    HMI_Message_Request : ARRAY[0..121] OF BOOL;  (* #HMI メッセージ表示要求; [0] 未使用; [1] 【Y616】A(左側) 供給スライド戻 異常表示; [2] 【Y617】A(左側) 供給スライド行 異常表示; [3] 【Y618】A(左側) 供給ピックアップ戻 異常表示; [4] 【Y619】A(左側) 供給ピックアップ行 異常表示; [5] 【Y620】A(左側) 供給チャック閉 戻 異常表示; [6] 【Y621】A(左側) 供給チャック開 行 異常表示; [7] 【Y622】B(右側) 供給スライド戻 異常表示; [8] 【Y623】B(右側) 供給スライド行 異常表示; [9] 【Y624】B(右側) 供給ピックアップ戻 異常表示; [10] 【Y625】B(右側) 供給ピックアップ行 異常表示; [11] 【Y626】B(右側) 供給チャック閉 戻 異常表示; [12] 【Y627】B(右側) 供給チャック開 行 異常表示; [13] 【Y700】A(左側) 高さ検査押え戻 異常表示; [14] 【Y701】A(左側) 高さ検査押え行 異常表示; [15] 【Y702】A(左側) 高さ検査持上戻 異常表示; [16] 【Y703】A(左側) 高さ検査持上行 異常表示; [17] 【Y704】A(左側) NG1ピックアップ戻 異常表示; [18] 【Y705】A(左側) NG1ピックアップ 行 異常表示; [19] 【Y706】A(左側) NG1チャック戻 異常表示; [20] 【Y707】A(左側) NG1チャック行 異常表示; [21] 【Y708】A(左側)ST4 反転1チャック閉 異常表示; [22] 【Y709】A(左側)ST4 反転1チャック開 異常表示; [23] 【Y710】A(左側)ST4 反転1ピックアップ戻 異常表示; [24] 【Y711】A(左側)ST4 反転1ピックアップ行 異常表示; [25] 【Y712】A(左側)ST6 反転2チャック閉 戻 異常表示; [26] 【Y713】A(左側)ST6 反転2チャック開 行 異常表示; [27] 【Y714】A(左側)ST6 反転2ピックアップ戻 異常表示; [28] 【Y715】A(左側)ST6 反転2ピックアップ行 異常表示; [29] 【Y716】A(左側) 排出チャック閉 戻 異常表示; [30] 【Y717】A(左側) 排出チャック開 行 異常表示; [31] 【Y718】A(左側) 排出フォルダ送り戻 異常表示; [32] 【Y719】A(左側) 排出フォルダ送り行 異常表示; [33] A(左側) 位置1ストッパー戻 異常表示; [34] 【Y720】A(左側) 位置1ストッパー 行 異常表示; [35] 【Y721】A(左側) 位置2ストッパー 異常表示; [36] 【Y721】A(左側) 位置2ストッパー 異常表示; [37] 【Y722】A(左側) 位置3ストッパー戻 異常表示; [38] 【Y722】A(左側) 位置3ストッパー行 異常表示; [39] Output_A_Error_M[33] 異常表示; [40] 【Y723】A(左側) 位置4ストッパー行 異常表示; [41] 【Y724】A(左側) 位置5ストッパー戻 異常表示; [42] 【Y724】A(左側) 位置5ストッパー行 異常表示; [43] 【Y725】A(左側) 位置6ストッパー戻 異常表示; [44] 【Y725】A(左側) 位置6ストッパー行 異常表示; [45] 【Y726】A(左側) ストックフォルダターン戻 異常表示; [46] 【Y727】A(左側) ストックフォルダターン行 異常表示; [47] 【Y728】A(左側) NG1仕分け 戻 異常表示; [48] 【Y729】A(左側) NG1仕分け 行 異常表示; [49] 【Y800】B(右側) 高さ検査押え戻 異常表示; [50] 【Y801】B(右側) 高さ検査押え行 異常表示; [51] 【Y802】B(右側) 高さ検査持上戻 異常表示; [52] 【Y803】B(右側) 高さ検査持上行 異常表示; [53] 【Y804】B(右側) NG1ピックアップ戻 異常表示; [54] 【Y805】B(右側) NG1ピックアップ 行 異常表示; [55] 【Y806】B(右側) NG1チャック戻 異常表示; [56] 【Y807】B(右側) NG1チャック行 異常表示; [57] 【Y808】B(右側)ST4 反転1チャック閉 戻 異常表示; [58] 【Y809】B(右側)ST4 反転1チャック開 戻 異常表示; [59] 【Y810】B(右側)ST4 反転1ピックアップ戻 異常表示; [60] 【Y811】B(右側)ST4 反転1ピックアップ行 異常表示; [61] 【Y812】B(右側)ST6 反転2チャック閉 戻 異常表示; [62] 【Y813】B(右側)ST6 反転2チャック開 行 異常表示; [63] 【Y814】B(右側)ST6 反転2ピックアップ戻 異常表示; [64] 【Y815】B(右側)ST6 反転2ピックアップ行 異常表示; [65] 【Y816】B(右側) 排出チャック閉 戻 異常表示; [66] 【Y817】B(右側) 排出チャック開 行 異常表示; [67] 【Y818】B(右側) 排出フォルダ送り戻 異常表示; [68] 【Y819】B(右側) 排出フォルダ送り行 異常表示; [69] 【Y820】B(右側) 位置1ストッパー 戻 異常表示; [70] 【Y820】B(右側) 位置1ストッパー 行 異常表示; [71] 【Y821】B(右側) 位置2ストッパー戻 異常表示; [72] 【Y821】B(右側) 位置2ストッパー行 異常表示; [73] 【Y822】B(右側) 位置3ストッパー戻 異常表示; [74] 【Y822】B(右側) 位置3ストッパー行 異常表示; [75] 【Y823】B(右側) 位置4ストッパー戻 異常表示; [76] 【Y823】B(右側) 位置4ストッパー行 異常表示; [77] 【Y824】B(右側) 位置5ストッパー戻 異常表示; [78] 【Y824】B(右側) 位置5ストッパー行 異常表示; [79] 【Y825】B(右側) 位置6ストッパー戻 異常表示; [80] 【Y825】B(右側) 位置6ストッパー行 異常表示; [81] 【Y826】B(右側) ストックフォルダターン戻 異常表示; [82] 【Y827】B(右側) ストックフォルダターン行 異常表示; [83] 【Y828】B(右側) NG1仕分け 戻 異常表示; [84] 【Y829】B(右側) NG1仕分け 行 異常表示; [85] 【Y1200】空コンテナ送り 戻 異常表示; [86] 【Y1201】空コンテナ送り 行 異常表示; [87] 【Y1202】段バラシ爪 戻 異常表示; [88] 【Y1203】段バラシ爪 行 異常表示; [89] 【Y1204】コンテナ排出 戻 異常表示; [90] 【Y1205】コンテナ排出 行 異常表示; [91] Output_Share_Error_M[7] 異常表示; [92] 【Y1207】箱入れチャック 行 異常表示; [93] 【Y1208】コンテナ仕分けストッパー 戻 異常表示; [94] 【Y1209】コンテナ仕分けストッパー 行 異常表示; [95] 【Y1210】コンテナ仕分け送り 戻 異常表示; [96] Output_Share_Error_M[12] 異常表示; [97] 【Y1300】A(左側) コンベア受渡送り戻 異常表示; [98] 【Y1301】A(左側) コンベア受渡送り行 異常表示; [99] 【Y1302】B(右側) コンベア受渡送り戻 異常表示; [100] 【Y1303】B(右側) コンベア受渡送り行 異常表示; [101] ST1 搬送ワーク不一致; [102] ST2 搬送ワーク不一致; [103] ST3 搬送ワーク不一致; [104] ST4 搬送ワーク不一致; [105] ST5 搬送ワーク不一致; [106] ST6 搬送ワーク不一致; [107] ST7 搬送ワーク不一致; [108] A(左側) ST1 FH測定時間超過; [109] A(左側) ST1 FH異常; [110] A(左側) ST5 FH異常; [111] B(右側) ST1 FH異常; [112] B(右側) ST5 FH異常; [113] A(左側) ST1 FH判定OK; [114] A(左側) ST1 FH判定NG1; [115] A(左側) ST1 FH判定NG2; [116] A(左側) ST1 検査前ワーク不一致; [117] A(左側) ST5 FH測定時間超過; [118] A(左側) ST5 FH判定OK; [119] A(左側) ST5 FH判定NG1; [120] A(左側) ST5 FH判定NG2; [121] A(左側) ST5 検査前ワーク不一致 *)
END_VAR

PROGRAM ModeManagement_モード管理
VAR
    Setting_M : BOOL;
    Manual_M : BOOL;
    Auto_M : BOOL;
    Dummy_M : BOOL;
    Inital_M : BOOL;
    Output_Error_M : ARRAY[0..99] OF Bool;
    Index_Error_001 : DINT;
    Index_B_001 : DINT;
    Index_Share_001 : DINT;
    Error_TON : ARRAY[0..99] OF TON;  (* [2] A(左側) ST1 測定タイムアウト; [4] A(左側) ST5 測定タイムアウト *)
    Error_TOF : ARRAY[0..99] OF TOF;
    AutoMode_A_M : ARRAY[0..99] OF Bool;
    ６ : DINT;
    ST4_A_Rev_01_Origin_M : ARRAY[0..99] OF Bool;  (* A(左側) ST4 反転1 原点復帰工程; [1] A(左側) ST4 反転1 原点復帰開始; [2] A(左側) ST4 反転1 原点復帰中; [3] A(左側) ST4 反転1 ピックアップ戻; [4] A(左側) ST4 反転1 モータ原点復帰開始; [5] A(左側) ST4 反転1 ピックアップ行; [6] A(左側) ST4 反転1 チャック閉; [7] A(左側) ST4 反転1 原点復帰完了（ワーク無） *)
    ST4_A_Rev_01_OriginDone : BOOL;  (* A(左側) ST4 反転1 原点復帰完了 *)
    ST4_A_Rev_02_Origin_M : ARRAY[0..99] OF Bool;  (* A(左側) ST6 反転2 原点復帰工程; [1] A(左側) ST6 反転2 原点復帰開始; [2] A(左側) ST6 反転2 原点復帰中; [3] A(左側) ST6 反転2 ピックアップ戻; [4] A(左側) ST6 反転2 モータ原点復帰開始; [5] A(左側) ST6 反転2 ピックアップ行; [6] A(左側) ST6 反転2 チャック閉; [7] A(左側) ST6 反転2 原点復帰完了（ワーク無） *)
    ST4_A_Rev_02_OriginDone : BOOL;  (* A(左側) ST6 反転2 原点復帰完了 *)
    ST4_B_Rev_01_Origin_M : ARRAY[0..99] OF Bool;  (* B(右側) ST4 反転1 原点復帰工程; [1] B(右側) ST4 反転1 原点復帰開始; [2] B(右側) ST4 反転1 原点復帰中; [3] B(右側) ST4 反転1 ピックアップ戻; [4] B(右側) ST4 反転1 モータ原点復帰開始; [5] B(右側) ST4 反転1 ピックアップ行; [6] B(右側) ST4 反転1 チャック閉; [7] B(右側) ST4 反転1 原点復帰完了（ワーク無） *)
    ST4_B_Rev_01_OriginDone : BOOL;  (* B(右側) ST4 反転1 原点復帰完了 *)
    ST4_B_Rev_02_Origin_M : ARRAY[0..99] OF Bool;  (* B(右側) ST6 反転2 原点復帰工程; [1] B(右側) ST6 反転2 原点復帰開始; [2] B(右側) ST6 反転2 原点復帰中; [3] B(右側) ST6 反転2 ピックアップ戻; [4] B(右側) ST6 反転2 モータ原点復帰開始; [5] B(右側) ST6 反転2 ピックアップ行; [6] B(右側) ST6 反転2 チャック閉; [7] B(右側) ST6 反転2 原点復帰完了（ワーク無） *)
    ST4_B_Rev_02_OriginDone : BOOL;  (* B(右側) ST6 反転2 原点復帰完了 *)
    Error_ST1_A_Timeout : BOOL;  (* FHタイムアウト（非保持） *)
    Error_ST5_A_Timeout : BOOL;  (* FHタイムアウト（非保持） *)
END_VAR
VAR_EXTERNAL
    Output_A_Error_M : ARRAY[0..99] OF Bool;
    Output_A_Restart_M : ARRAY[0..99] OF Bool;
    In_Sw_RESET : BOOL;
    In_Sw_START : BOOL;
    ManualMode : BOOL;
    M9999 : BOOL;
    Output_B_Error_M : ARRAY[0..99] OF Bool;  (* B(右側)シリンダエラー *)
    Output_B_Restart_M : ARRAY[0..99] OF Bool;  (* B(右側)シリンダ再開： *)
    Output_Share_Error_M : ARRAY[0..99] OF Bool;
    Output_Share_Restart_M : ARRAY[0..99] OF Bool;
    TimerQ_In_Sen_Accum_CV_A_Full : BOOL;
    Out_TDC_Stop : BOOL;
    In_Sen_Unl_Conv_A_Pass : BOOL;
    In_Sen_Accum_CV_A_Full : BOOL;
    In_Sen_Unl_Conv_B_Pass : BOOL;
    Pause : ARRAY[0..99] OF Bool;  (* [3] FH A(左側) ST1; [9] FH A(左側) ST5; [10] FH B(右側) ST1; [11] FH B(右側) ST5; [12] A(左側) ST6 反転2 ワーク不一致 *)
    AutoMode : BOOL;
    In_Sen_DOOR_01 : BOOL;
    In_Sen_DOOR_02 : BOOL;
    In_Sen_DOOR_03 : BOOL;
    In_Sen_DOOR_04 : BOOL;
    In_Sen_DOOR_05 : BOOL;
    In_Sen_DOOR_06 : BOOL;
    In_Sw_EMS1 : BOOL;
    In_Sw_EMS2 : BOOL;
    In_Sw_EMS3 : BOOL;
    In_Sen_AIR１_Pressure_01 : BOOL;
    In_Sen_AIR１_Pressure_02 : BOOL;
    In_Sen_AIR１_Pressure_03 : BOOL;
    TEST_M : ARRAY[0..99] OF Bool;
    ST0_Sup_Start : BOOL;  (* ST0_動作開始 *)
    Out_CYw_Sply_Pick_A_H_Auto : ARRAY[0..10] OF Bool;
    Out_CYw_Sply_Pick_A_H_Done : BOOL;
    Out_CYw_Sply_Slide_A_H_Auto : ARRAY[0..10] OF Bool;
    Out_CYw_Sply_Slide_A_H_Done : BOOL;
    Out_CYw_Sup_Chuck_A_Cl_H_Auto : ARRAY[0..10] OF Bool;
    Out_CYw_Sup_Chuck_A_Cl_H_Done : BOOL;
    In_Sen_Accum_CV_A_Arrival : BOOL;
    In_Sen_Work_A_Pos_00 : BOOL;
    Out_CYw_Sply_Pick_A_F_Auto : ARRAY[0..10] OF Bool;
    Out_CYw_Sply_Pick_A_F_Done : BOOL;
    Out_CYw_Sup_Chuck_A_Cl_F_Auto : ARRAY[0..10] OF Bool;
    Out_CYw_Sup_Chuck_A_Cl_F_Done : BOOL;
    Out_CYw_Sply_Slide_A_F_Auto : ARRAY[0..10] OF Bool;
    Out_CYw_Sply_Slide_A_F_Done : BOOL;
    Ins_A_Cv_Error : BOOL;
    Station_A_Data : ARRAY[0..8] OF sData;
    Ins_A_Cv_M : ARRAY[0..99] OF Bool;
    HMI_MessageNo : ARRAY[0..9] OF UINT;
    FH_5552_10_A_Auto : BOOL;
    In_Sen_Accum_CV_B_Full : BOOL;
    FH_Line3_Error_Status_1 : BOOL;
    FH_Line0_Error_Status_1 : BOOL;
    FH_Line1_Error_Status_1 : BOOL;
    FH_Line2_Error_Status_1 : BOOL;
    FH_Line0_Error_Clear_1 : BOOL;
    FH_Line1_Error_Clear_1 : BOOL;
    FH_Line2_Error_Clear_1 : BOOL;
    FH_Line3_Error_Clear_1 : BOOL;
    Ins_A_Next_Cycle : BOOL;
    OriginDone : BOOL;  (* 原点復帰完了 *)
    DummyDone : BOOL;  (* ダミーチェック完了 *)
    HMI_CurrentPage : STRING[256];
    Ins_A_End : BOOL;
    Auto_A_Start : BOOL;  (* 自動運転 開始 *)
    Auto_Ready : BOOL;  (* 自動運転可能 *)
    ST0_A_Sup_Busy : BOOL;
    ST1_A_Ca1_Busy : BOOL;
    RCON1_1_IN_Alarm : BOOL;  (* 軸異常 *)
    RCON1_1_IN_EmergencyStop : BOOL;  (* 非常停止状態（監視） *)
    RCON1_1_Error : BOOL;  (* 異常予備（未接続） *)
    RCON1_1_IN_HomeDone : BOOL;  (* 原点復帰完了 *)
    RCON1_1_Error_Clear : BOOL;  (* 解除予備（未接続） *)
    Error_M : ARRAY[0..99] OF Bool;  (* エラー：; [1] シリンダ; [2] コンベア＆ドアセンサ; [3] 未使用：Error_ST1_A_M[0]へ移行; [4] A(左側)検査コンベア ワーク不一致; [5] 未使用：Error_ST3_A_M[1]へ移行; [9] 未使用：Error_ST5_A_M[0]へ移行; [10] 未使用：Error_ST1_B_M[0]へ移行; [11] 未使用：Error_ST5_B_M[0]へ移行; [12] 未使用：Error_ST6_A_M[0]へ移行 *)
    ST1_A_Ca1_M : ARRAY[0..99] OF Bool;  (* [6] A(左側) ST1 検査前ワーク不一致 *)
    ST2_A_Hgt_M : ARRAY[0..99] OF Bool;
    ST3_A_Dis1_M : ARRAY[0..99] OF Bool;
    HMI_Home_SW : BOOL;
    Origin_Busy : BOOL;  (* 原点復帰中 *)
    Out_CYw_Rev_01_Pick_A_H_Origin : ARRAY[0..10] OF Bool;  (* 原点復帰【Y710】A(左側)ST4 反転1ピックアップ戻： *)
    Out_CYw_Rev_01_Pick_A_H_Done : BOOL;  (* 【Y710】A(左側)ST4 反転1ピックアップ戻 動作完了 *)
    Stm_A_Rev_Axis000_Origin : BOOL;  (* A(左側) ST4 反転1 モータ原点復帰開始 *)
    Stm_A_Rev_Axis000_OriginDone : BOOL;  (* A(左側) ST4 反転1 モータ原点復帰完了 *)
    Out_CYw_Rev_01_Pick_A_F_Origin : ARRAY[0..99] OF Bool;  (* 原点復帰【Y711】A(左側)ST4 反転1ピックアップ行： *)
    Out_CYw_Rev_01_Pick_A_F_Done : BOOL;  (* 【Y711】A(左側)ST4 反転1ピックアップ行 動作完了 *)
    Out_CYw_Rev_01_Chk_A_H_Origin : ARRAY[0..99] OF Bool;  (* 原点復帰【Y708】A(左側)ST4 反転1チャック閉： *)
    Out_CYw_Rev_01_Chk_A_H_Done : BOOL;  (* 【Y708】A(左側)ST4 反転1チャック閉 動作完了 *)
    TimerQ_In_Sen_Work_A_Pos_04 : BOOL;
    Out_CYw_Rev_02_Pick_A_H_Origin : ARRAY[0..10] OF Bool;  (* 原点復帰 【Y714】A(左側)ST6 反転2ピックアップ戻 *)
    Out_CYw_Rev_02_Pick_A_H_Done : BOOL;  (* 【Y714】A(左側)ST6 反転2ピックアップ戻 動作完了 *)
    Stm_A_Rev_Axis001_Origin : BOOL;  (* A(左側) ST6 反転2 モータ原点復帰開始 *)
    Stm_A_Rev_Axis001_OriginDone : BOOL;  (* A(左側) ST6 反転2 モータ原点復帰完了 *)
    Out_CYw_Rev_02_Pick_A_F_Origin : ARRAY[0..99] OF Bool;  (* 原点復帰 【Y715】A(左側)ST6 反転2ピックアップ行 *)
    Out_CYw_Rev_02_Pick_A_F_Done : BOOL;  (* 【Y715】A(左側)ST6 反転2ピックアップ行 動作完了 *)
    Out_CYw_Rev_02_Chk_A_H_Origin : ARRAY[0..99] OF Bool;  (* 原点復帰 【Y712】A(左側)ST6 反転2チャック閉 戻 *)
    Out_CYw_Rev_02_Chk_A_H_Done : BOOL;  (* 【Y712】A(左側)ST6 反転2チャック閉 戻 動作完了 *)
    TimerQ_In_Sen_Work_A_Pos_06 : BOOL;  (* 【X208】A(左側)ワーク位置6 *)
    Auto_B_Start : BOOL;  (* B(右側)自動運転開始（後続処理未接続） *)
    Out_CYw_Rev_01_Pick_B_H_Origin : ARRAY[0..10] OF Bool;  (* 原点復帰 【Y810】B(右側)ST4 反転1ピックアップ戻 *)
    Out_CYw_Rev_01_Pick_B_H_Done : BOOL;  (* 【Y810】B(右側)ST4 反転1ピックアップ戻 動作完了 *)
    Stm_B_Rev_Axis002_Origin : BOOL;  (* B(右側) ST4 反転1 モータ原点復帰開始 *)
    Stm_B_Rev_Axis002_OriginDone : BOOL;  (* B(右側) ST4 反転1 モータ原点復帰完了 *)
    Out_CYw_Rev_01_Pick_B_F_Origin : ARRAY[0..99] OF Bool;  (* 原点復帰 【Y811】B(右側)ST4 反転1ピックアップ行 *)
    Out_CYw_Rev_01_Pick_B_F_Done : BOOL;  (* 【Y811】B(右側)ST4 反転1ピックアップ行 動作完了 *)
    Out_CYw_Rev_01_Chk_B_H_Origin : ARRAY[0..99] OF Bool;  (* 原点復帰 【Y808】B(右側)ST4 反転1チャック閉 戻 *)
    Out_CYw_Rev_01_Chk_B_H_Done : BOOL;  (* 【Y808】B(右側)ST4 反転1チャック閉 戻 動作完了 *)
    TimerQ_In_Sen_Work_B_Pos_04 : BOOL;  (* 【X406】B(右側)ワーク位置4 *)
    Out_CYw_Rev_02_Pick_B_H_Origin : ARRAY[0..10] OF Bool;  (* 原点復帰 【Y814】B(右側)ST6 反転2ピックアップ戻 *)
    Out_CYw_Rev_02_Pick_B_H_Done : BOOL;  (* 【Y814】B(右側)ST6 反転2ピックアップ戻 動作完了 *)
    Stm_B_Rev_Axis003_Origin : BOOL;  (* B(右側) ST6 反転2 モータ原点復帰開始 *)
    Stm_B_Rev_Axis003_OriginDone : BOOL;  (* B(右側) ST6 反転2 モータ原点復帰完了 *)
    Out_CYw_Rev_02_Pick_B_F_Origin : ARRAY[0..99] OF Bool;  (* 原点復帰 【Y815】B(右側)ST6 反転2ピックアップ行 *)
    Out_CYw_Rev_02_Pick_B_F_Done : BOOL;  (* 【Y815】B(右側)ST6 反転2ピックアップ行 動作完了 *)
    Out_CYw_Rev_02_Chk_B_H_Origin : ARRAY[0..99] OF Bool;  (* 原点復帰 【Y812】B(右側)ST6 反転2チャック閉 戻 *)
    Out_CYw_Rev_02_Chk_B_H_Done : BOOL;  (* 【Y812】B(右側)ST6 反転2チャック閉 戻 動作完了 *)
    TimerQ_In_Sen_Work_B_Pos_06 : BOOL;  (* 【X408】B(右側)ワーク位置6 *)
    ST4_A_Rev1_M : ARRAY[0..99] OF Bool;  (* [10] A(左側) ST4 ワーク不一致エラー; [12] 【Y708】A(左側) ST4 反転1チャック閉 *)
    ST5_A_Ca2_M : ARRAY[0..99] OF Bool;  (* A(左側) ST5 カメラ2工程; [1] A(左側) ST5 カメラ2検査開始; [2] 【Y724】A(左側) ST5 ストッパー戻; [3] A(左側) ST5 ワーク有無判定; [4] A(左側) ST5 ワーク有; [5] A(左側) ST5 ワーク無; [6] A(左側) ST5 検査前ワーク不一致; [7] A(左側) ST5 FH測定開始 *)
    FH_A_ST5_Auto : BOOL;  (* A(左側) ST5 FH自動測定 *)
END_VAR
VAR_EXTERNAL CONSTANT
    ST6_A_Rev2_M : ARRAY[0..99] OF Bool;  (* A(左側) ST6 反転2工程; [1] A(左側) ST6 反転2 動作開始; [2] A(左側) ST6 反転2 【Y714】ピックアップ戻; [3] A(左側) ST6 反転2 【Y725】位置6ストッパー戻; [4] A(左側) ST6 反転2 原点角度転送; [5] A(左側) ST6 反転2 原点位置移動開始; [6] A(左側) ST6 反転2 原点位置移動完了; [7] A(左側) ST6 反転2 ワーク有無判定; [8] A(左側) ST6 反転2 ワーク有・前工程OK; [9] A(左側) ST6 反転2 ワーク無・前工程NG; [10] A(左側) ST6 反転2 ワーク不一致エラー; [11] A(左側) ST6 反転2 【Y715】反転前ピックアップ行; [12] A(左側) ST6 反転2 【Y712】チャック閉; [13] A(左側) ST6 反転2 【Y714】反転前ピックアップ戻; [14] A(左側) ST6 反転2 反転角度転送; [15] A(左側) ST6 反転2 反転位置移動完了; [16] A(左側) ST6 反転2 【Y715】設置ピックアップ行; [17] A(左側) ST6 反転2 【Y713】チャック開; [18] A(左側) ST6 反転2 【Y714】設置ピックアップ戻 *)
END_VAR
VAR_EXTERNAL
    ST7_A_Dis2_M : ARRAY[0..99] OF Bool;  (* [9] ST7 A ワーク有; [10] ST3 A ワーク無; [11] ST7 排出前ワーク不一致エラー; [12] コンベア下降 位置転送; [13] コンベア下降 移動開始; [14] 排出チャック開 行; [15] セイフティ上昇 位置転送; [16] セイフティ上昇 移動開始; [17] NG / フォルダストック 仕分け IAI移動位置 判定; [18] ストックフォルダ位置; [19] カメラ2 キズNG位置; [20] カメラ2 姿NG位置; [21] 排出フォルダ送り行; [22] SF/NG2左右 移動開始; [23] SF/NG2上下 目標位置転送; [24] ストックフォルダ カウントup; [25] カメラ キズNG位置; [26] カメラ 姿NG位置; [27] SF/NG2上下 移動開始; [28] 排出チャック戻／ワーク解放; [29] SF/NG2上下 原点位置転送; [30] SF/NG2上下 原点移動開始; [31] SF/NG2左右 原点位置転送; [32] 排出フォルダ送り戻; [33] 排出フォルダ戻完了 *)
    Error_ST1_A_M : ARRAY[0..4] OF BOOL;  (* #A(左側) ST1 カメラ1 異常; [0] 総合異常; [1] 機器異常; [2] タイムアウト; [3] ワーク不一致; [4] 予備（監視なし） *)
    Error_ST1_B_M : ARRAY[0..4] OF BOOL;  (* #B(右側) ST1 カメラ1 異常; [0] 総合異常; [1] 機器異常; [2] 予備（監視なし）; [3] 予備（監視なし）; [4] 予備（監視なし） *)
    Error_ST2_A_M : ARRAY[0..4] OF BOOL;  (* #A(左側) ST2 高さ検査 異常; [0] 総合異常; [1] 予備（監視なし）; [2] 予備（監視なし）; [3] ワーク不一致; [4] 予備（監視なし） *)
    Error_ST3_A_M : ARRAY[0..4] OF BOOL;  (* #A(左側) ST3 NG1排出 異常; [0] 総合異常; [1] 機器異常; [2] 予備（監視なし）; [3] ワーク不一致; [4] 予備（監視なし） *)
    Error_ST4_A_M : ARRAY[0..4] OF BOOL;  (* #A(左側) ST4 反転1 異常; [0] 総合異常; [1] 予備（監視なし）; [2] 予備（監視なし）; [3] ワーク不一致; [4] 予備（監視なし） *)
    Error_ST5_A_M : ARRAY[0..4] OF BOOL;  (* #A(左側) ST5 カメラ2 異常; [0] 総合異常; [1] 機器異常; [2] タイムアウト; [3] ワーク不一致; [4] 予備（監視なし） *)
    Error_ST5_B_M : ARRAY[0..4] OF BOOL;  (* #B(右側) ST5 カメラ2 異常; [0] 総合異常; [1] 機器異常; [2] 予備（監視なし）; [3] 予備（監視なし）; [4] 予備（監視なし） *)
    Error_ST6_A_M : ARRAY[0..4] OF BOOL;  (* #A(左側) ST6 反転2 異常; [0] 総合異常; [1] 予備（監視なし）; [2] 予備（監視なし）; [3] ワーク不一致; [4] 予備（監視なし） *)
    Error_ST7_A_M : ARRAY[0..4] OF BOOL;  (* #A(左側) ST7 SF排出 異常; [0] 総合異常; [1] 予備（監視なし）; [2] 予備（監視なし）; [3] ワーク不一致; [4] 満杯 *)
    Error_ST7_A_Source_M : ARRAY[0..4] OF BOOL;  (* #A(左側) ST7 発生理由（内部保持）; [3] ワーク不一致; [4] 満杯（既存B側入力） *)
    HMI_Message_Request : ARRAY[0..121] OF BOOL;  (* #HMI メッセージ表示要求; [0] 未使用; [1] 【Y616】A(左側) 供給スライド戻 異常表示; [2] 【Y617】A(左側) 供給スライド行 異常表示; [3] 【Y618】A(左側) 供給ピックアップ戻 異常表示; [4] 【Y619】A(左側) 供給ピックアップ行 異常表示; [5] 【Y620】A(左側) 供給チャック閉 戻 異常表示; [6] 【Y621】A(左側) 供給チャック開 行 異常表示; [7] 【Y622】B(右側) 供給スライド戻 異常表示; [8] 【Y623】B(右側) 供給スライド行 異常表示; [9] 【Y624】B(右側) 供給ピックアップ戻 異常表示; [10] 【Y625】B(右側) 供給ピックアップ行 異常表示; [11] 【Y626】B(右側) 供給チャック閉 戻 異常表示; [12] 【Y627】B(右側) 供給チャック開 行 異常表示; [13] 【Y700】A(左側) 高さ検査押え戻 異常表示; [14] 【Y701】A(左側) 高さ検査押え行 異常表示; [15] 【Y702】A(左側) 高さ検査持上戻 異常表示; [16] 【Y703】A(左側) 高さ検査持上行 異常表示; [17] 【Y704】A(左側) NG1ピックアップ戻 異常表示; [18] 【Y705】A(左側) NG1ピックアップ 行 異常表示; [19] 【Y706】A(左側) NG1チャック戻 異常表示; [20] 【Y707】A(左側) NG1チャック行 異常表示; [21] 【Y708】A(左側)ST4 反転1チャック閉 異常表示; [22] 【Y709】A(左側)ST4 反転1チャック開 異常表示; [23] 【Y710】A(左側)ST4 反転1ピックアップ戻 異常表示; [24] 【Y711】A(左側)ST4 反転1ピックアップ行 異常表示; [25] 【Y712】A(左側)ST6 反転2チャック閉 戻 異常表示; [26] 【Y713】A(左側)ST6 反転2チャック開 行 異常表示; [27] 【Y714】A(左側)ST6 反転2ピックアップ戻 異常表示; [28] 【Y715】A(左側)ST6 反転2ピックアップ行 異常表示; [29] 【Y716】A(左側) 排出チャック閉 戻 異常表示; [30] 【Y717】A(左側) 排出チャック開 行 異常表示; [31] 【Y718】A(左側) 排出フォルダ送り戻 異常表示; [32] 【Y719】A(左側) 排出フォルダ送り行 異常表示; [33] A(左側) 位置1ストッパー戻 異常表示; [34] 【Y720】A(左側) 位置1ストッパー 行 異常表示; [35] 【Y721】A(左側) 位置2ストッパー 異常表示; [36] 【Y721】A(左側) 位置2ストッパー 異常表示; [37] 【Y722】A(左側) 位置3ストッパー戻 異常表示; [38] 【Y722】A(左側) 位置3ストッパー行 異常表示; [39] Output_A_Error_M[33] 異常表示; [40] 【Y723】A(左側) 位置4ストッパー行 異常表示; [41] 【Y724】A(左側) 位置5ストッパー戻 異常表示; [42] 【Y724】A(左側) 位置5ストッパー行 異常表示; [43] 【Y725】A(左側) 位置6ストッパー戻 異常表示; [44] 【Y725】A(左側) 位置6ストッパー行 異常表示; [45] 【Y726】A(左側) ストックフォルダターン戻 異常表示; [46] 【Y727】A(左側) ストックフォルダターン行 異常表示; [47] 【Y728】A(左側) NG1仕分け 戻 異常表示; [48] 【Y729】A(左側) NG1仕分け 行 異常表示; [49] 【Y800】B(右側) 高さ検査押え戻 異常表示; [50] 【Y801】B(右側) 高さ検査押え行 異常表示; [51] 【Y802】B(右側) 高さ検査持上戻 異常表示; [52] 【Y803】B(右側) 高さ検査持上行 異常表示; [53] 【Y804】B(右側) NG1ピックアップ戻 異常表示; [54] 【Y805】B(右側) NG1ピックアップ 行 異常表示; [55] 【Y806】B(右側) NG1チャック戻 異常表示; [56] 【Y807】B(右側) NG1チャック行 異常表示; [57] 【Y808】B(右側)ST4 反転1チャック閉 戻 異常表示; [58] 【Y809】B(右側)ST4 反転1チャック開 戻 異常表示; [59] 【Y810】B(右側)ST4 反転1ピックアップ戻 異常表示; [60] 【Y811】B(右側)ST4 反転1ピックアップ行 異常表示; [61] 【Y812】B(右側)ST6 反転2チャック閉 戻 異常表示; [62] 【Y813】B(右側)ST6 反転2チャック開 行 異常表示; [63] 【Y814】B(右側)ST6 反転2ピックアップ戻 異常表示; [64] 【Y815】B(右側)ST6 反転2ピックアップ行 異常表示; [65] 【Y816】B(右側) 排出チャック閉 戻 異常表示; [66] 【Y817】B(右側) 排出チャック開 行 異常表示; [67] 【Y818】B(右側) 排出フォルダ送り戻 異常表示; [68] 【Y819】B(右側) 排出フォルダ送り行 異常表示; [69] 【Y820】B(右側) 位置1ストッパー 戻 異常表示; [70] 【Y820】B(右側) 位置1ストッパー 行 異常表示; [71] 【Y821】B(右側) 位置2ストッパー戻 異常表示; [72] 【Y821】B(右側) 位置2ストッパー行 異常表示; [73] 【Y822】B(右側) 位置3ストッパー戻 異常表示; [74] 【Y822】B(右側) 位置3ストッパー行 異常表示; [75] 【Y823】B(右側) 位置4ストッパー戻 異常表示; [76] 【Y823】B(右側) 位置4ストッパー行 異常表示; [77] 【Y824】B(右側) 位置5ストッパー戻 異常表示; [78] 【Y824】B(右側) 位置5ストッパー行 異常表示; [79] 【Y825】B(右側) 位置6ストッパー戻 異常表示; [80] 【Y825】B(右側) 位置6ストッパー行 異常表示; [81] 【Y826】B(右側) ストックフォルダターン戻 異常表示; [82] 【Y827】B(右側) ストックフォルダターン行 異常表示; [83] 【Y828】B(右側) NG1仕分け 戻 異常表示; [84] 【Y829】B(右側) NG1仕分け 行 異常表示; [85] 【Y1200】空コンテナ送り 戻 異常表示; [86] 【Y1201】空コンテナ送り 行 異常表示; [87] 【Y1202】段バラシ爪 戻 異常表示; [88] 【Y1203】段バラシ爪 行 異常表示; [89] 【Y1204】コンテナ排出 戻 異常表示; [90] 【Y1205】コンテナ排出 行 異常表示; [91] Output_Share_Error_M[7] 異常表示; [92] 【Y1207】箱入れチャック 行 異常表示; [93] 【Y1208】コンテナ仕分けストッパー 戻 異常表示; [94] 【Y1209】コンテナ仕分けストッパー 行 異常表示; [95] 【Y1210】コンテナ仕分け送り 戻 異常表示; [96] Output_Share_Error_M[12] 異常表示; [97] 【Y1300】A(左側) コンベア受渡送り戻 異常表示; [98] 【Y1301】A(左側) コンベア受渡送り行 異常表示; [99] 【Y1302】B(右側) コンベア受渡送り戻 異常表示; [100] 【Y1303】B(右側) コンベア受渡送り行 異常表示; [101] ST1 搬送ワーク不一致; [102] ST2 搬送ワーク不一致; [103] ST3 搬送ワーク不一致; [104] ST4 搬送ワーク不一致; [105] ST5 搬送ワーク不一致; [106] ST6 搬送ワーク不一致; [107] ST7 搬送ワーク不一致; [108] A(左側) ST1 FH測定時間超過; [109] A(左側) ST1 FH異常; [110] A(左側) ST5 FH異常; [111] B(右側) ST1 FH異常; [112] B(右側) ST5 FH異常; [113] A(左側) ST1 FH判定OK; [114] A(左側) ST1 FH判定NG1; [115] A(左側) ST1 FH判定NG2; [116] A(左側) ST1 検査前ワーク不一致; [117] A(左側) ST5 FH測定時間超過; [118] A(左側) ST5 FH判定OK; [119] A(左側) ST5 FH判定NG1; [120] A(左側) ST5 FH判定NG2; [121] A(左側) ST5 検査前ワーク不一致 *)
END_VAR
VAR
    _p1 : BOOL;
    _p2 : BOOL;
    _p3 : BOOL;
    _p4 : BOOL;
    _p5 : BOOL;
    _p6 : BOOL;
    _p7 : BOOL;
    _p8 : BOOL;
    _p9 : BOOL;
    _p10 : BOOL;
    _p11 : BOOL;
    _p12 : BOOL;
    _p13 : BOOL;
    _p14 : BOOL;
    _p15 : BOOL;
    _p16 : BOOL;
    _p17 : BOOL;
    _p18 : BOOL;
    _p19 : BOOL;
    _p20 : BOOL;
    _p21 : BOOL;
    _p22 : BOOL;
    _p23 : BOOL;
    _p24 : BOOL;
    _e25 : R_TRIG;
    _e26 : R_TRIG;
    _e27 : R_TRIG;
    _e28 : R_TRIG;
    _e29 : R_TRIG;
    _e30 : R_TRIG;
    _e31 : R_TRIG;
    _e32 : R_TRIG;
    _e33 : R_TRIG;
    _p34 : BOOL;
    _p35 : BOOL;
    _p36 : BOOL;
    _p37 : BOOL;
    _e38 : R_TRIG;
    _e39 : R_TRIG;
    _e40 : R_TRIG;
    _e41 : R_TRIG;
    _e42 : R_TRIG;
    _e43 : R_TRIG;
    _e44 : R_TRIG;
    _e45 : R_TRIG;
    _p46 : BOOL;
END_VAR

(* Section Initial_初期化処理: ladder, written here as Structured Text *)

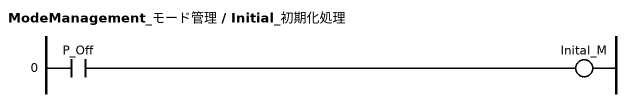
(* Rung 0 *)
Inital_M := P_Off;

(* Section Origin_原点復帰: ladder, written here as Structured Text *)

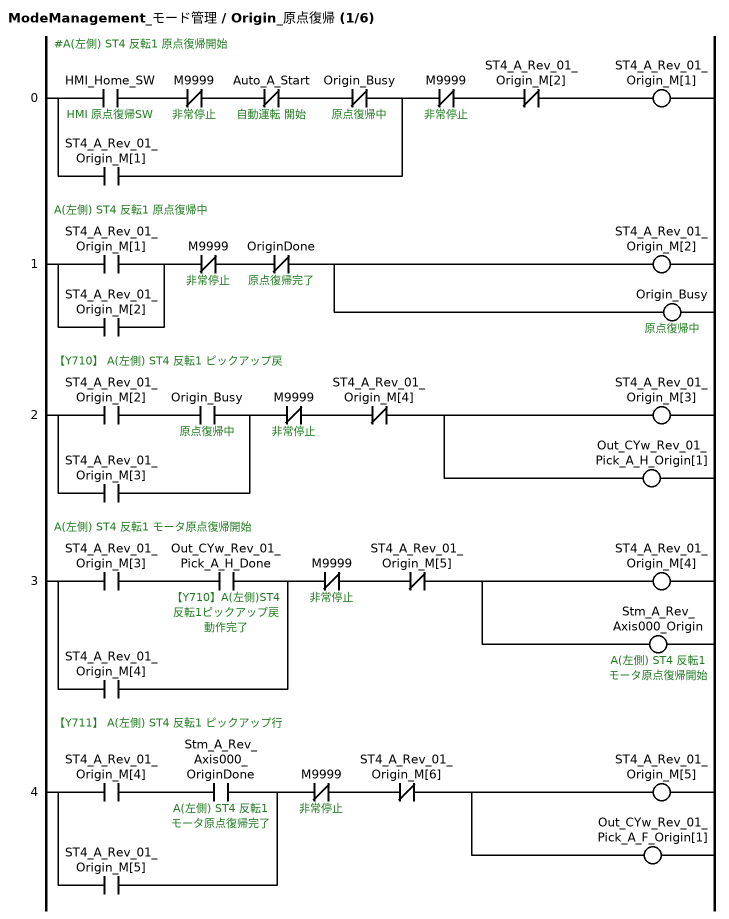
(* Rung 0: #A(左側) ST4 反転1 原点復帰開始 *)
ST4_A_Rev_01_Origin_M[1] := ((HMI_Home_SW AND NOT M9999 AND NOT Auto_A_Start AND NOT Origin_Busy) OR ST4_A_Rev_01_Origin_M[1]) AND NOT M9999 AND NOT ST4_A_Rev_01_Origin_M[2];
(* Rung 1: A(左側) ST4 反転1 原点復帰中 *)
_p1 := (ST4_A_Rev_01_Origin_M[1] OR ST4_A_Rev_01_Origin_M[2]) AND NOT M9999 AND NOT OriginDone;
ST4_A_Rev_01_Origin_M[2] := _p1;
Origin_Busy := _p1;
(* Rung 2: 【Y710】 A(左側) ST4 反転1 ピックアップ戻 *)
_p2 := ((ST4_A_Rev_01_Origin_M[2] AND Origin_Busy) OR ST4_A_Rev_01_Origin_M[3]) AND NOT M9999 AND NOT ST4_A_Rev_01_Origin_M[4];
ST4_A_Rev_01_Origin_M[3] := _p2;
Out_CYw_Rev_01_Pick_A_H_Origin[1] := _p2;
(* Rung 3: A(左側) ST4 反転1 モータ原点復帰開始 *)
_p3 := ((ST4_A_Rev_01_Origin_M[3] AND Out_CYw_Rev_01_Pick_A_H_Done) OR ST4_A_Rev_01_Origin_M[4]) AND NOT M9999 AND NOT ST4_A_Rev_01_Origin_M[5];
ST4_A_Rev_01_Origin_M[4] := _p3;
Stm_A_Rev_Axis000_Origin := _p3;
(* Rung 4: 【Y711】 A(左側) ST4 反転1 ピックアップ行 *)
_p4 := ((ST4_A_Rev_01_Origin_M[4] AND Stm_A_Rev_Axis000_OriginDone) OR ST4_A_Rev_01_Origin_M[5]) AND NOT M9999 AND NOT ST4_A_Rev_01_Origin_M[6];
ST4_A_Rev_01_Origin_M[5] := _p4;
Out_CYw_Rev_01_Pick_A_F_Origin[1] := _p4;

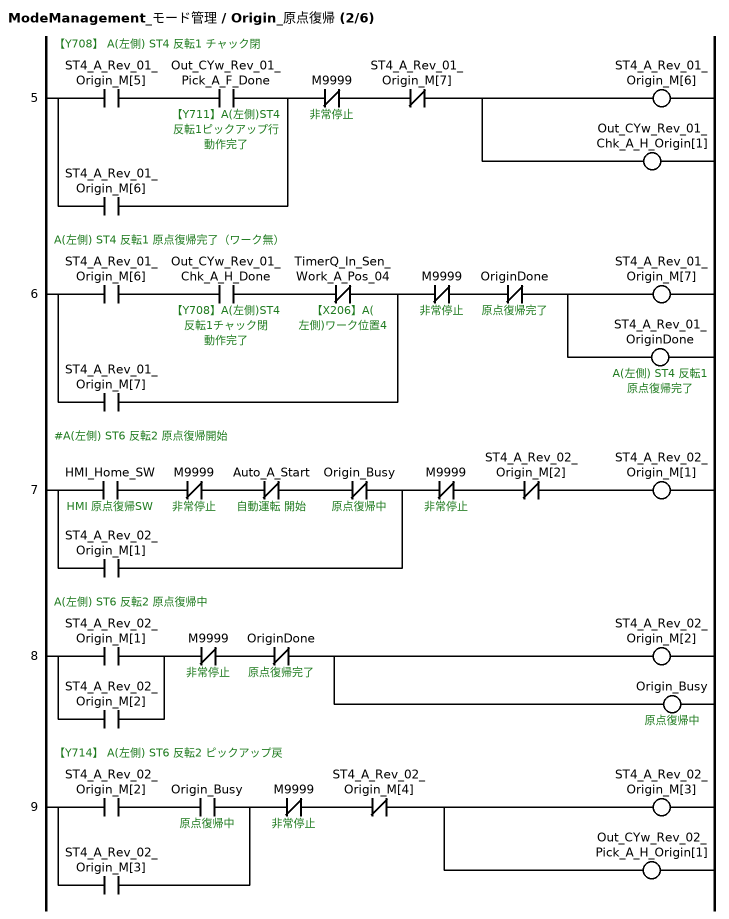
(* Rung 5: 【Y708】 A(左側) ST4 反転1 チャック閉 *)
_p5 := ((ST4_A_Rev_01_Origin_M[5] AND Out_CYw_Rev_01_Pick_A_F_Done) OR ST4_A_Rev_01_Origin_M[6]) AND NOT M9999 AND NOT ST4_A_Rev_01_Origin_M[7];
ST4_A_Rev_01_Origin_M[6] := _p5;
Out_CYw_Rev_01_Chk_A_H_Origin[1] := _p5;
(* Rung 6: A(左側) ST4 反転1 原点復帰完了（ワーク無） *)
_p6 := ((ST4_A_Rev_01_Origin_M[6] AND Out_CYw_Rev_01_Chk_A_H_Done AND NOT TimerQ_In_Sen_Work_A_Pos_04) OR ST4_A_Rev_01_Origin_M[7]) AND NOT M9999 AND NOT OriginDone;
ST4_A_Rev_01_Origin_M[7] := _p6;
ST4_A_Rev_01_OriginDone := _p6;
(* Rung 7: #A(左側) ST6 反転2 原点復帰開始 *)
ST4_A_Rev_02_Origin_M[1] := ((HMI_Home_SW AND NOT M9999 AND NOT Auto_A_Start AND NOT Origin_Busy) OR ST4_A_Rev_02_Origin_M[1]) AND NOT M9999 AND NOT ST4_A_Rev_02_Origin_M[2];
(* Rung 8: A(左側) ST6 反転2 原点復帰中 *)
_p7 := (ST4_A_Rev_02_Origin_M[1] OR ST4_A_Rev_02_Origin_M[2]) AND NOT M9999 AND NOT OriginDone;
ST4_A_Rev_02_Origin_M[2] := _p7;
Origin_Busy := _p7;
(* Rung 9: 【Y714】 A(左側) ST6 反転2 ピックアップ戻 *)
_p8 := ((ST4_A_Rev_02_Origin_M[2] AND Origin_Busy) OR ST4_A_Rev_02_Origin_M[3]) AND NOT M9999 AND NOT ST4_A_Rev_02_Origin_M[4];
ST4_A_Rev_02_Origin_M[3] := _p8;
Out_CYw_Rev_02_Pick_A_H_Origin[1] := _p8;

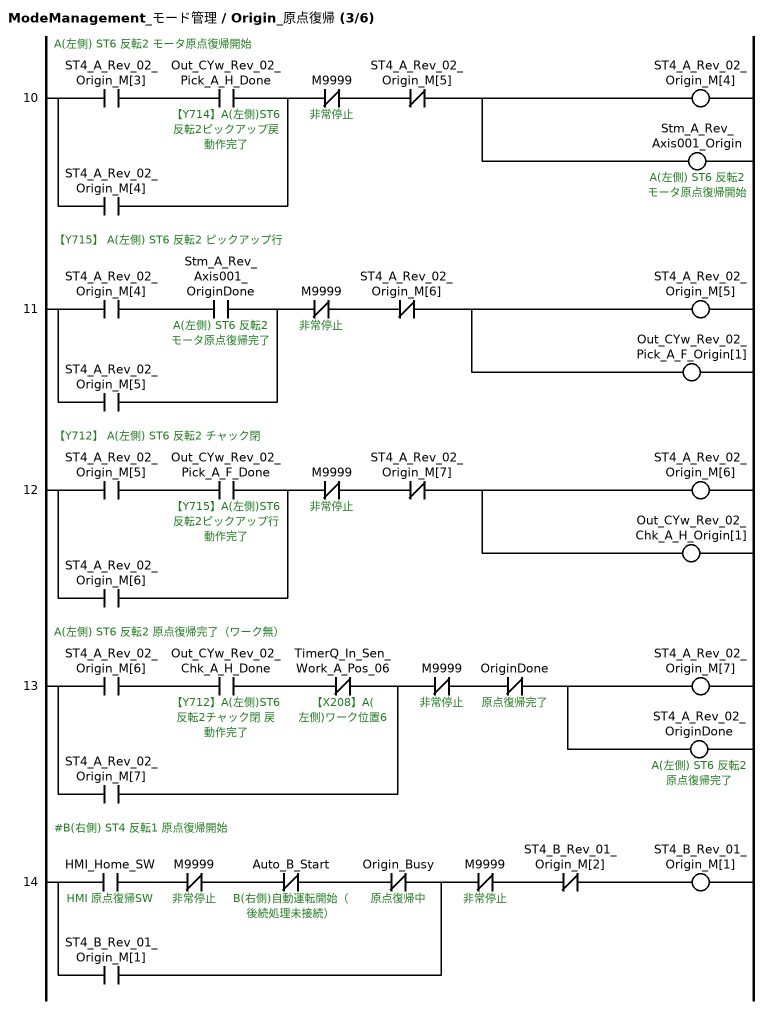
(* Rung 10: A(左側) ST6 反転2 モータ原点復帰開始 *)
_p9 := ((ST4_A_Rev_02_Origin_M[3] AND Out_CYw_Rev_02_Pick_A_H_Done) OR ST4_A_Rev_02_Origin_M[4]) AND NOT M9999 AND NOT ST4_A_Rev_02_Origin_M[5];
ST4_A_Rev_02_Origin_M[4] := _p9;
Stm_A_Rev_Axis001_Origin := _p9;
(* Rung 11: 【Y715】 A(左側) ST6 反転2 ピックアップ行 *)
_p10 := ((ST4_A_Rev_02_Origin_M[4] AND Stm_A_Rev_Axis001_OriginDone) OR ST4_A_Rev_02_Origin_M[5]) AND NOT M9999 AND NOT ST4_A_Rev_02_Origin_M[6];
ST4_A_Rev_02_Origin_M[5] := _p10;
Out_CYw_Rev_02_Pick_A_F_Origin[1] := _p10;
(* Rung 12: 【Y712】 A(左側) ST6 反転2 チャック閉 *)
_p11 := ((ST4_A_Rev_02_Origin_M[5] AND Out_CYw_Rev_02_Pick_A_F_Done) OR ST4_A_Rev_02_Origin_M[6]) AND NOT M9999 AND NOT ST4_A_Rev_02_Origin_M[7];
ST4_A_Rev_02_Origin_M[6] := _p11;
Out_CYw_Rev_02_Chk_A_H_Origin[1] := _p11;
(* Rung 13: A(左側) ST6 反転2 原点復帰完了（ワーク無） *)
_p12 := ((ST4_A_Rev_02_Origin_M[6] AND Out_CYw_Rev_02_Chk_A_H_Done AND NOT TimerQ_In_Sen_Work_A_Pos_06) OR ST4_A_Rev_02_Origin_M[7]) AND NOT M9999 AND NOT OriginDone;
ST4_A_Rev_02_Origin_M[7] := _p12;
ST4_A_Rev_02_OriginDone := _p12;
(* Rung 14: #B(右側) ST4 反転1 原点復帰開始 *)
ST4_B_Rev_01_Origin_M[1] := ((HMI_Home_SW AND NOT M9999 AND NOT Auto_B_Start AND NOT Origin_Busy) OR ST4_B_Rev_01_Origin_M[1]) AND NOT M9999 AND NOT ST4_B_Rev_01_Origin_M[2];

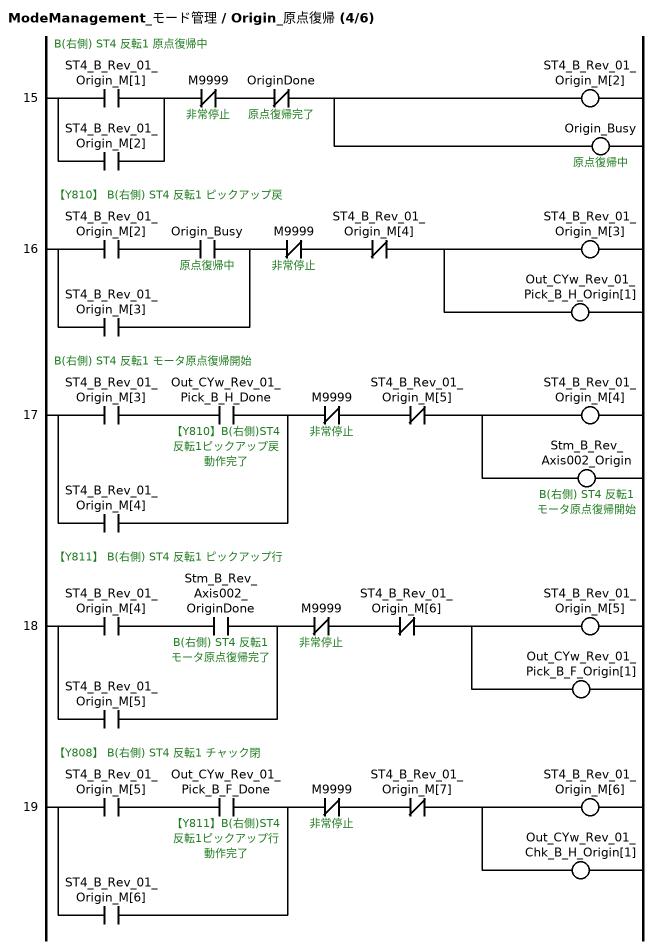
(* Rung 15: B(右側) ST4 反転1 原点復帰中 *)
_p13 := (ST4_B_Rev_01_Origin_M[1] OR ST4_B_Rev_01_Origin_M[2]) AND NOT M9999 AND NOT OriginDone;
ST4_B_Rev_01_Origin_M[2] := _p13;
Origin_Busy := _p13;
(* Rung 16: 【Y810】 B(右側) ST4 反転1 ピックアップ戻 *)
_p14 := ((ST4_B_Rev_01_Origin_M[2] AND Origin_Busy) OR ST4_B_Rev_01_Origin_M[3]) AND NOT M9999 AND NOT ST4_B_Rev_01_Origin_M[4];
ST4_B_Rev_01_Origin_M[3] := _p14;
Out_CYw_Rev_01_Pick_B_H_Origin[1] := _p14;
(* Rung 17: B(右側) ST4 反転1 モータ原点復帰開始 *)
_p15 := ((ST4_B_Rev_01_Origin_M[3] AND Out_CYw_Rev_01_Pick_B_H_Done) OR ST4_B_Rev_01_Origin_M[4]) AND NOT M9999 AND NOT ST4_B_Rev_01_Origin_M[5];
ST4_B_Rev_01_Origin_M[4] := _p15;
Stm_B_Rev_Axis002_Origin := _p15;
(* Rung 18: 【Y811】 B(右側) ST4 反転1 ピックアップ行 *)
_p16 := ((ST4_B_Rev_01_Origin_M[4] AND Stm_B_Rev_Axis002_OriginDone) OR ST4_B_Rev_01_Origin_M[5]) AND NOT M9999 AND NOT ST4_B_Rev_01_Origin_M[6];
ST4_B_Rev_01_Origin_M[5] := _p16;
Out_CYw_Rev_01_Pick_B_F_Origin[1] := _p16;
(* Rung 19: 【Y808】 B(右側) ST4 反転1 チャック閉 *)
_p17 := ((ST4_B_Rev_01_Origin_M[5] AND Out_CYw_Rev_01_Pick_B_F_Done) OR ST4_B_Rev_01_Origin_M[6]) AND NOT M9999 AND NOT ST4_B_Rev_01_Origin_M[7];
ST4_B_Rev_01_Origin_M[6] := _p17;
Out_CYw_Rev_01_Chk_B_H_Origin[1] := _p17;

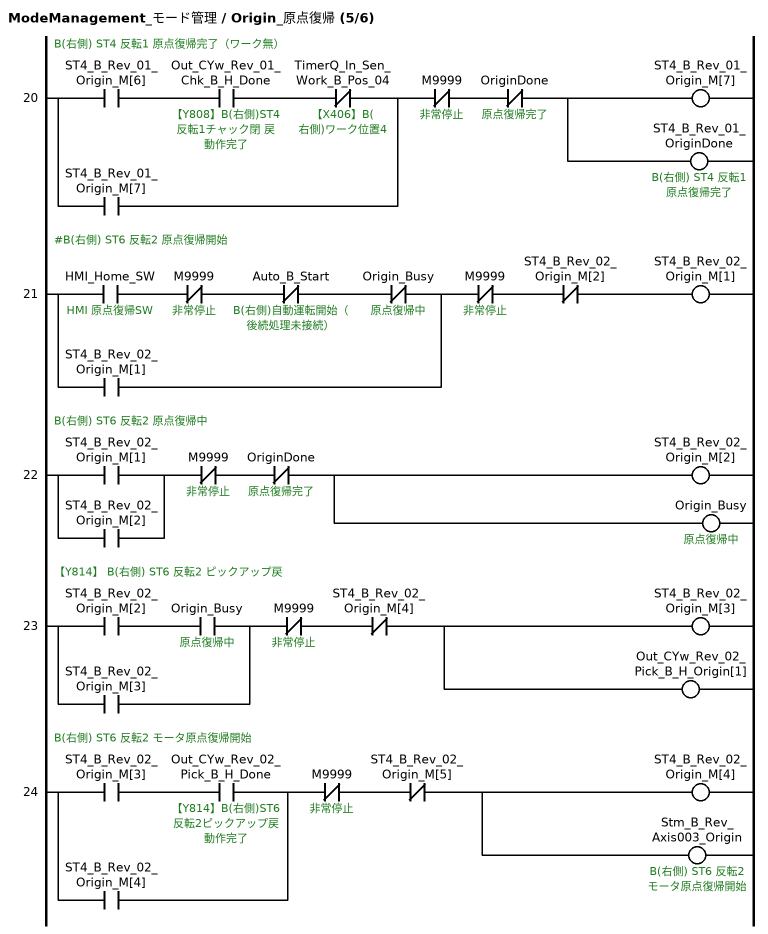
(* Rung 20: B(右側) ST4 反転1 原点復帰完了（ワーク無） *)
_p18 := ((ST4_B_Rev_01_Origin_M[6] AND Out_CYw_Rev_01_Chk_B_H_Done AND NOT TimerQ_In_Sen_Work_B_Pos_04) OR ST4_B_Rev_01_Origin_M[7]) AND NOT M9999 AND NOT OriginDone;
ST4_B_Rev_01_Origin_M[7] := _p18;
ST4_B_Rev_01_OriginDone := _p18;
(* Rung 21: #B(右側) ST6 反転2 原点復帰開始 *)
ST4_B_Rev_02_Origin_M[1] := ((HMI_Home_SW AND NOT M9999 AND NOT Auto_B_Start AND NOT Origin_Busy) OR ST4_B_Rev_02_Origin_M[1]) AND NOT M9999 AND NOT ST4_B_Rev_02_Origin_M[2];
(* Rung 22: B(右側) ST6 反転2 原点復帰中 *)
_p19 := (ST4_B_Rev_02_Origin_M[1] OR ST4_B_Rev_02_Origin_M[2]) AND NOT M9999 AND NOT OriginDone;
ST4_B_Rev_02_Origin_M[2] := _p19;
Origin_Busy := _p19;
(* Rung 23: 【Y814】 B(右側) ST6 反転2 ピックアップ戻 *)
_p20 := ((ST4_B_Rev_02_Origin_M[2] AND Origin_Busy) OR ST4_B_Rev_02_Origin_M[3]) AND NOT M9999 AND NOT ST4_B_Rev_02_Origin_M[4];
ST4_B_Rev_02_Origin_M[3] := _p20;
Out_CYw_Rev_02_Pick_B_H_Origin[1] := _p20;
(* Rung 24: B(右側) ST6 反転2 モータ原点復帰開始 *)
_p21 := ((ST4_B_Rev_02_Origin_M[3] AND Out_CYw_Rev_02_Pick_B_H_Done) OR ST4_B_Rev_02_Origin_M[4]) AND NOT M9999 AND NOT ST4_B_Rev_02_Origin_M[5];
ST4_B_Rev_02_Origin_M[4] := _p21;
Stm_B_Rev_Axis003_Origin := _p21;

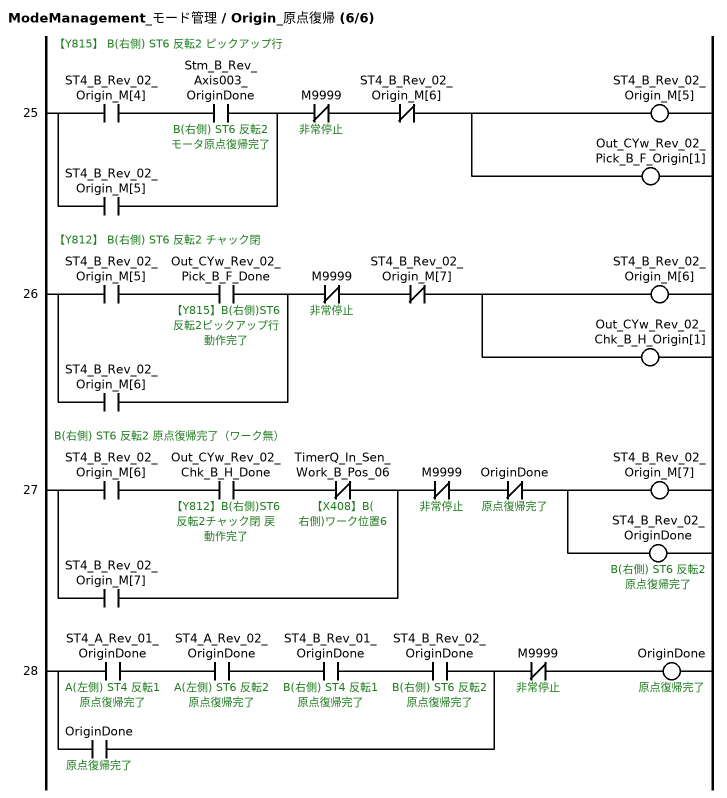
(* Rung 25: 【Y815】 B(右側) ST6 反転2 ピックアップ行 *)
_p22 := ((ST4_B_Rev_02_Origin_M[4] AND Stm_B_Rev_Axis003_OriginDone) OR ST4_B_Rev_02_Origin_M[5]) AND NOT M9999 AND NOT ST4_B_Rev_02_Origin_M[6];
ST4_B_Rev_02_Origin_M[5] := _p22;
Out_CYw_Rev_02_Pick_B_F_Origin[1] := _p22;
(* Rung 26: 【Y812】 B(右側) ST6 反転2 チャック閉 *)
_p23 := ((ST4_B_Rev_02_Origin_M[5] AND Out_CYw_Rev_02_Pick_B_F_Done) OR ST4_B_Rev_02_Origin_M[6]) AND NOT M9999 AND NOT ST4_B_Rev_02_Origin_M[7];
ST4_B_Rev_02_Origin_M[6] := _p23;
Out_CYw_Rev_02_Chk_B_H_Origin[1] := _p23;
(* Rung 27: B(右側) ST6 反転2 原点復帰完了（ワーク無） *)
_p24 := ((ST4_B_Rev_02_Origin_M[6] AND Out_CYw_Rev_02_Chk_B_H_Done AND NOT TimerQ_In_Sen_Work_B_Pos_06) OR ST4_B_Rev_02_Origin_M[7]) AND NOT M9999 AND NOT OriginDone;
ST4_B_Rev_02_Origin_M[7] := _p24;
ST4_B_Rev_02_OriginDone := _p24;
(* Rung 28 *)
OriginDone := ((ST4_A_Rev_01_OriginDone AND ST4_A_Rev_02_OriginDone AND ST4_B_Rev_01_OriginDone AND ST4_B_Rev_02_OriginDone) OR OriginDone) AND NOT M9999;

(* Section DummyCheck_ダミーチェック: ladder, written here as Structured Text *)

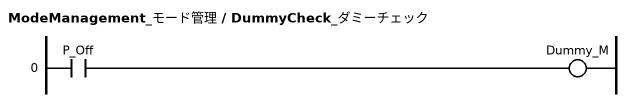
(* Rung 0 *)
Dummy_M := P_Off;

(* Section AutoMode_自動運転: ladder, written here as Structured Text *)

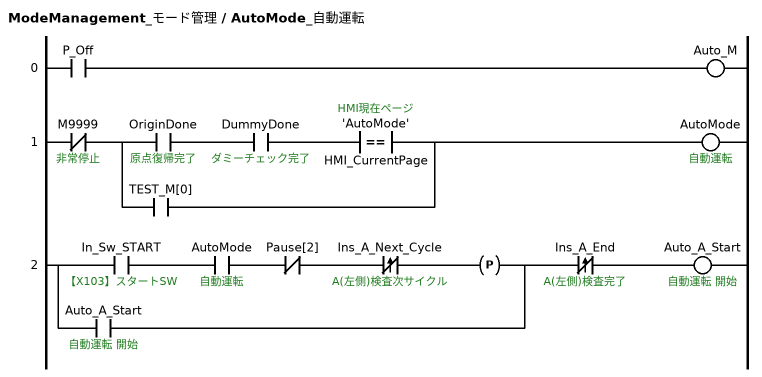
(* Rung 0 *)
Auto_M := P_Off;
(* Rung 1 *)
AutoMode := NOT M9999 AND ((OriginDone AND DummyDone AND ('AutoMode' = HMI_CurrentPage)) OR TEST_M[0]);
(* Rung 2 *)
_e25(CLK := Ins_A_Next_Cycle);
_e26(CLK := In_Sw_START AND AutoMode AND NOT Pause[2] AND NOT _e25.Q);
_e27(CLK := Ins_A_End);
Auto_A_Start := (_e26.Q OR Auto_A_Start) AND NOT _e27.Q;

(* Section Manual_手動運転: ladder, written here as Structured Text *)

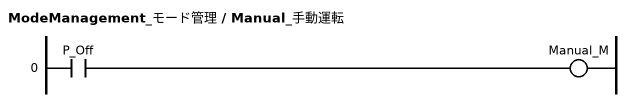
(* Rung 0 *)
Manual_M := P_Off;

(* Section Setting_設定: ladder, written here as Structured Text *)

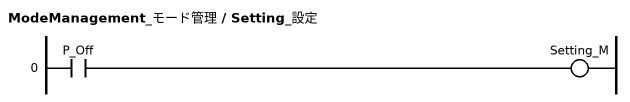
(* Rung 0 *)
Setting_M := P_Off;

(* Section Error_エラー処理: ladder, written here as Structured Text *)

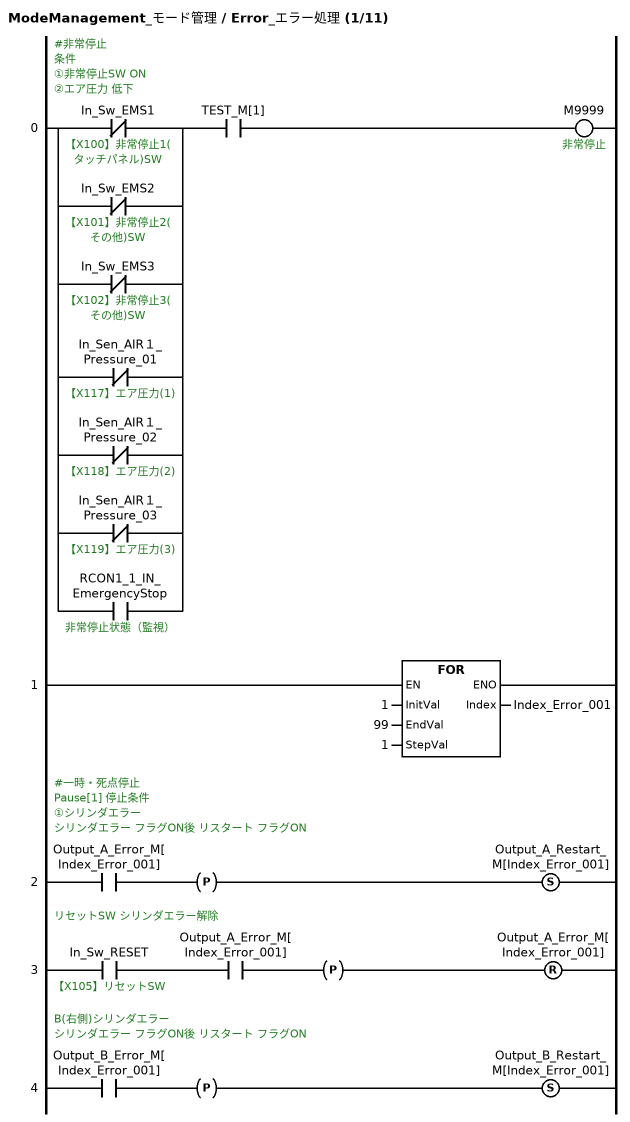
(* Rung 0: #非常停止 / 条件 / ①非常停止SW ON / ②エア圧力 低下 *)
M9999 := (NOT In_Sw_EMS1 OR NOT In_Sw_EMS2 OR NOT In_Sw_EMS3 OR NOT In_Sen_AIR１_Pressure_01 OR NOT In_Sen_AIR１_Pressure_02 OR NOT In_Sen_AIR１_Pressure_03 OR RCON1_1_IN_EmergencyStop) AND TEST_M[1];
(* Rung 1 *)
Index_Error_001 := FOR(InitVal := 1, EndVal := 99, StepVal := 1);
(* Rung 2: #一時・死点停止 / Pause[1] 停止条件 / ①シリンダエラー / シリンダエラー フラグON後 リスタート フラグON *)
_e28(CLK := Output_A_Error_M[Index_Error_001]);
IF _e28.Q THEN Output_A_Restart_M[Index_Error_001] := TRUE; END_IF;
(* Rung 3: リセットSW シリンダエラー解除 *)
_e29(CLK := In_Sw_RESET AND Output_A_Error_M[Index_Error_001]);
IF _e29.Q THEN Output_A_Error_M[Index_Error_001] := FALSE; END_IF;
(* Rung 4: B(右側)シリンダエラー / シリンダエラー フラグON後 リスタート フラグON *)
_e30(CLK := Output_B_Error_M[Index_Error_001]);
IF _e30.Q THEN Output_B_Restart_M[Index_Error_001] := TRUE; END_IF;

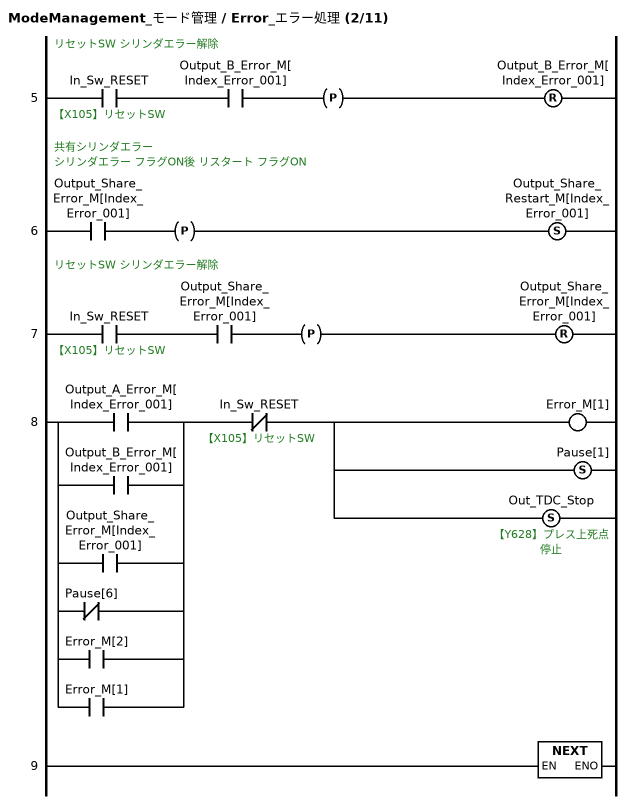
(* Rung 5: リセットSW シリンダエラー解除 *)
_e31(CLK := In_Sw_RESET AND Output_B_Error_M[Index_Error_001]);
IF _e31.Q THEN Output_B_Error_M[Index_Error_001] := FALSE; END_IF;
(* Rung 6: 共有シリンダエラー / シリンダエラー フラグON後 リスタート フラグON *)
_e32(CLK := Output_Share_Error_M[Index_Error_001]);
IF _e32.Q THEN Output_Share_Restart_M[Index_Error_001] := TRUE; END_IF;
(* Rung 7: リセットSW シリンダエラー解除 *)
_e33(CLK := In_Sw_RESET AND Output_Share_Error_M[Index_Error_001]);
IF _e33.Q THEN Output_Share_Error_M[Index_Error_001] := FALSE; END_IF;
(* Rung 8 *)
_p34 := (Output_A_Error_M[Index_Error_001] OR Output_B_Error_M[Index_Error_001] OR Output_Share_Error_M[Index_Error_001] OR NOT Pause[6] OR Error_M[2] OR Error_M[1]) AND NOT In_Sw_RESET;
Error_M[1] := _p34;
IF _p34 THEN
    Pause[1] := TRUE;
    Out_TDC_Stop := TRUE;
END_IF;
(* Rung 9 *)
NEXT();

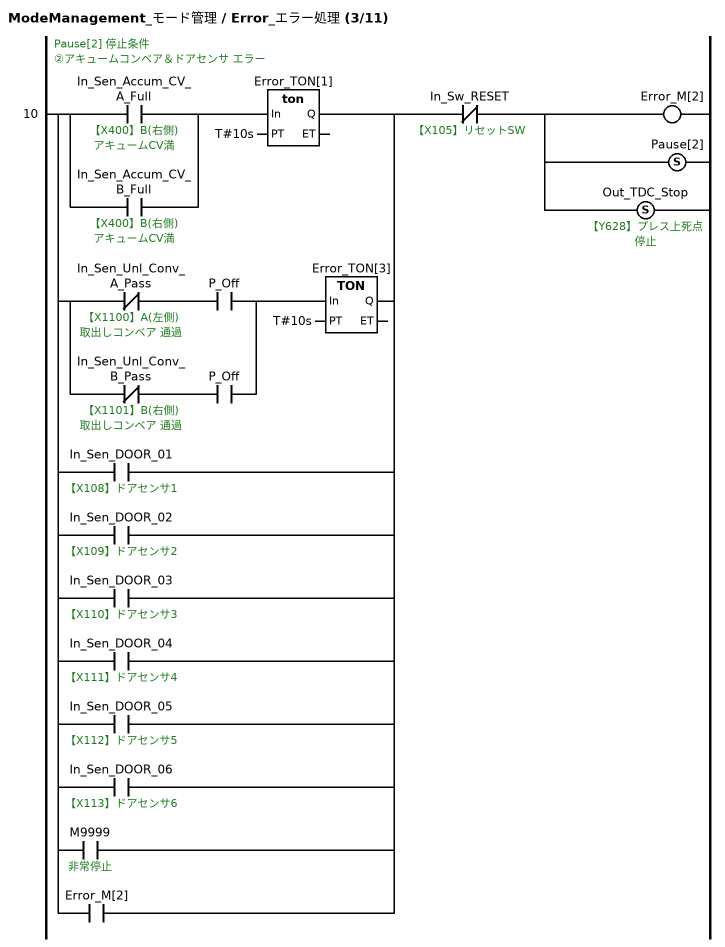
(* Rung 10: Pause[2] 停止条件 / ②アキュームコンベア＆ドアセンサ エラー *)
Error_TON[1](In := In_Sen_Accum_CV_A_Full OR In_Sen_Accum_CV_B_Full, PT := T#10s);
_p35 := Error_TON[1].Q;
Error_TON[3](In := (NOT In_Sen_Unl_Conv_A_Pass AND P_Off) OR (NOT In_Sen_Unl_Conv_B_Pass AND P_Off), PT := T#10s);
_p36 := (_p35 OR Error_TON[3].Q OR In_Sen_DOOR_01 OR In_Sen_DOOR_02 OR In_Sen_DOOR_03 OR In_Sen_DOOR_04 OR In_Sen_DOOR_05 OR In_Sen_DOOR_06 OR M9999 OR Error_M[2]) AND NOT In_Sw_RESET;
Error_M[2] := _p36;
IF _p36 THEN
    Pause[2] := TRUE;
    Out_TDC_Stop := TRUE;
END_IF;

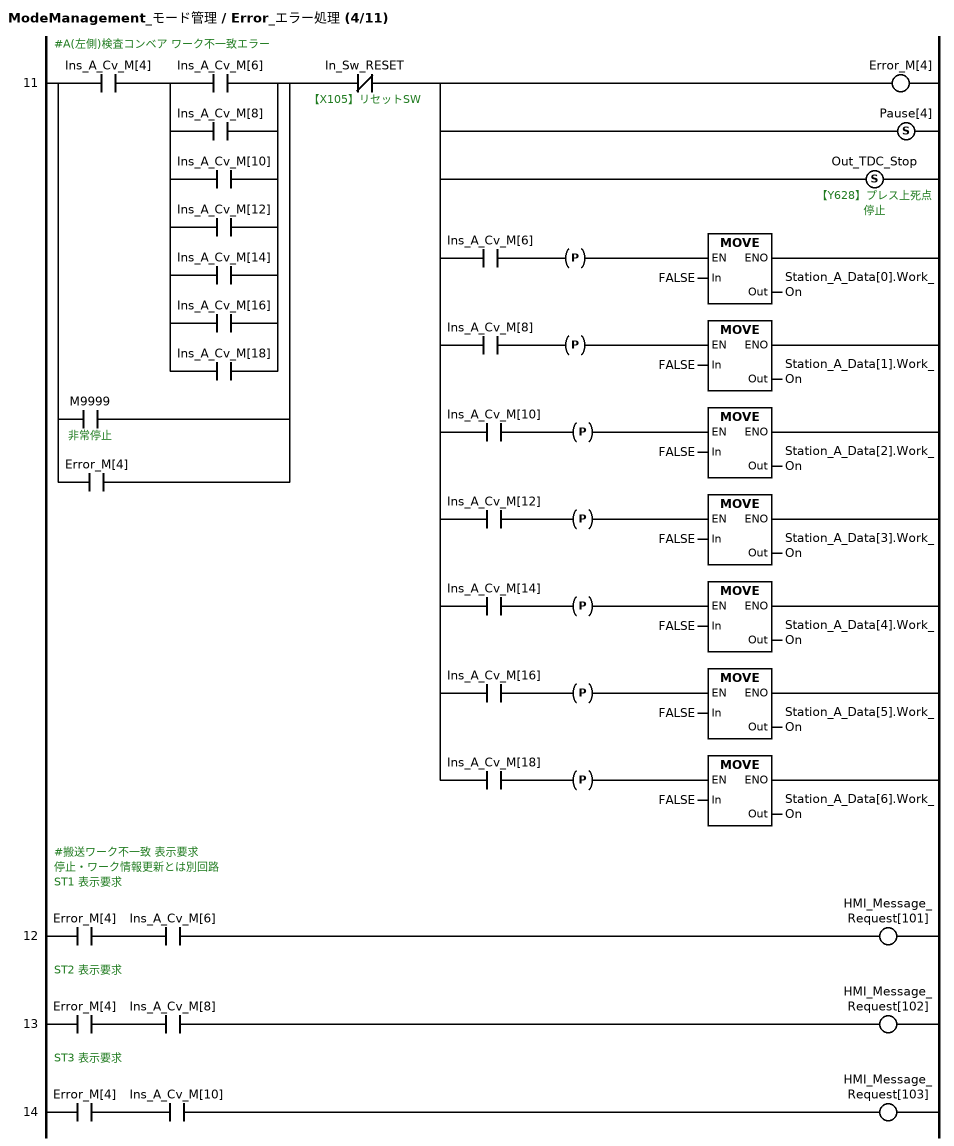
(* Rung 11: #A(左側)検査コンベア ワーク不一致エラー *)
_p37 := ((Ins_A_Cv_M[4] AND (Ins_A_Cv_M[6] OR Ins_A_Cv_M[8] OR Ins_A_Cv_M[10] OR Ins_A_Cv_M[12] OR Ins_A_Cv_M[14] OR Ins_A_Cv_M[16] OR Ins_A_Cv_M[18])) OR M9999 OR Error_M[4]) AND NOT In_Sw_RESET;
Error_M[4] := _p37;
IF _p37 THEN
    Pause[4] := TRUE;
    Out_TDC_Stop := TRUE;
END_IF;
_e38(CLK := _p37 AND Ins_A_Cv_M[6]);
IF _e38.Q THEN Station_A_Data[0].Work_On := FALSE; END_IF;
_e39(CLK := _p37 AND Ins_A_Cv_M[8]);
IF _e39.Q THEN Station_A_Data[1].Work_On := FALSE; END_IF;
_e40(CLK := _p37 AND Ins_A_Cv_M[10]);
IF _e40.Q THEN Station_A_Data[2].Work_On := FALSE; END_IF;
_e41(CLK := _p37 AND Ins_A_Cv_M[12]);
IF _e41.Q THEN Station_A_Data[3].Work_On := FALSE; END_IF;
_e42(CLK := _p37 AND Ins_A_Cv_M[14]);
IF _e42.Q THEN Station_A_Data[4].Work_On := FALSE; END_IF;
_e43(CLK := _p37 AND Ins_A_Cv_M[16]);
IF _e43.Q THEN Station_A_Data[5].Work_On := FALSE; END_IF;
_e44(CLK := _p37 AND Ins_A_Cv_M[18]);
IF _e44.Q THEN Station_A_Data[6].Work_On := FALSE; END_IF;
(* Rung 12: #搬送ワーク不一致 表示要求 / 停止・ワーク情報更新とは別回路 / ST1 表示要求 *)
HMI_Message_Request[101] := Error_M[4] AND Ins_A_Cv_M[6];
(* Rung 13: ST2 表示要求 *)
HMI_Message_Request[102] := Error_M[4] AND Ins_A_Cv_M[8];
(* Rung 14: ST3 表示要求 *)
HMI_Message_Request[103] := Error_M[4] AND Ins_A_Cv_M[10];

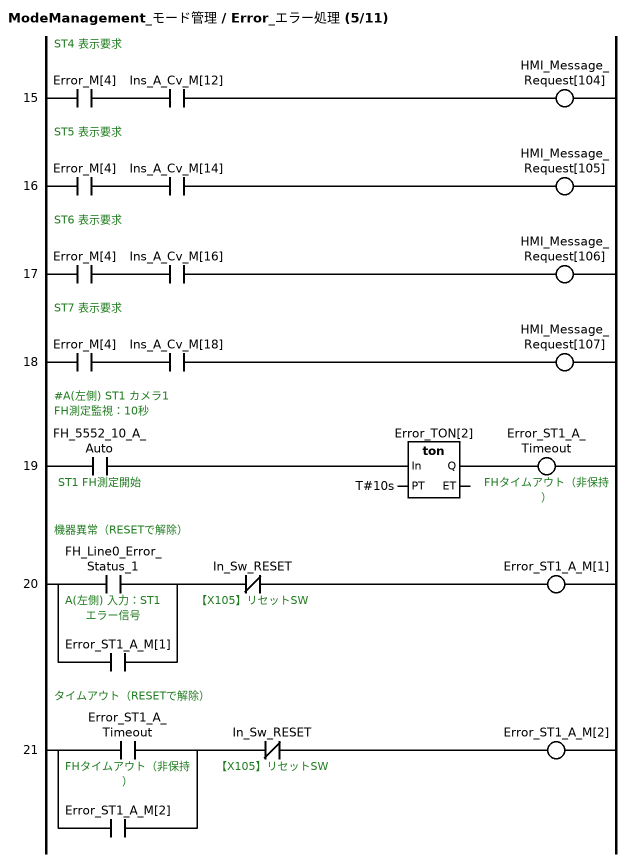
(* Rung 15: ST4 表示要求 *)
HMI_Message_Request[104] := Error_M[4] AND Ins_A_Cv_M[12];
(* Rung 16: ST5 表示要求 *)
HMI_Message_Request[105] := Error_M[4] AND Ins_A_Cv_M[14];
(* Rung 17: ST6 表示要求 *)
HMI_Message_Request[106] := Error_M[4] AND Ins_A_Cv_M[16];
(* Rung 18: ST7 表示要求 *)
HMI_Message_Request[107] := Error_M[4] AND Ins_A_Cv_M[18];
(* Rung 19: #A(左側) ST1 カメラ1 / FH測定監視：10秒 *)
Error_TON[2](In := FH_5552_10_A_Auto, PT := T#10s);
Error_ST1_A_Timeout := Error_TON[2].Q;
(* Rung 20: 機器異常（RESETで解除） *)
Error_ST1_A_M[1] := (FH_Line0_Error_Status_1 OR Error_ST1_A_M[1]) AND NOT In_Sw_RESET;
(* Rung 21: タイムアウト（RESETで解除） *)
Error_ST1_A_M[2] := (Error_ST1_A_Timeout OR Error_ST1_A_M[2]) AND NOT In_Sw_RESET;

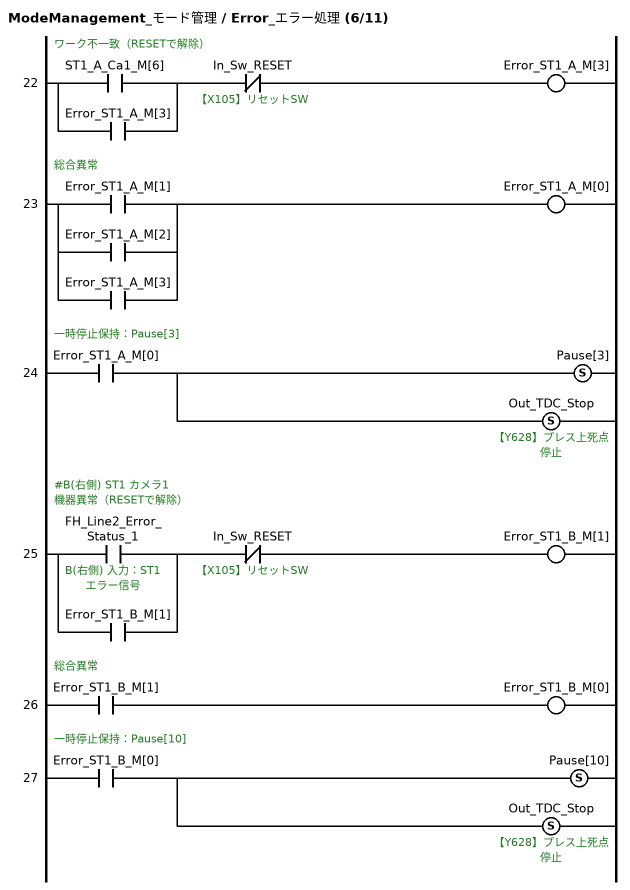
(* Rung 22: ワーク不一致（RESETで解除） *)
Error_ST1_A_M[3] := (ST1_A_Ca1_M[6] OR Error_ST1_A_M[3]) AND NOT In_Sw_RESET;
(* Rung 23: 総合異常 *)
Error_ST1_A_M[0] := Error_ST1_A_M[1] OR Error_ST1_A_M[2] OR Error_ST1_A_M[3];
(* Rung 24: 一時停止保持：Pause[3] *)
IF Error_ST1_A_M[0] THEN
    Pause[3] := TRUE;
    Out_TDC_Stop := TRUE;
END_IF;
(* Rung 25: #B(右側) ST1 カメラ1 / 機器異常（RESETで解除） *)
Error_ST1_B_M[1] := (FH_Line2_Error_Status_1 OR Error_ST1_B_M[1]) AND NOT In_Sw_RESET;
(* Rung 26: 総合異常 *)
Error_ST1_B_M[0] := Error_ST1_B_M[1];
(* Rung 27: 一時停止保持：Pause[10] *)
IF Error_ST1_B_M[0] THEN
    Pause[10] := TRUE;
    Out_TDC_Stop := TRUE;
END_IF;

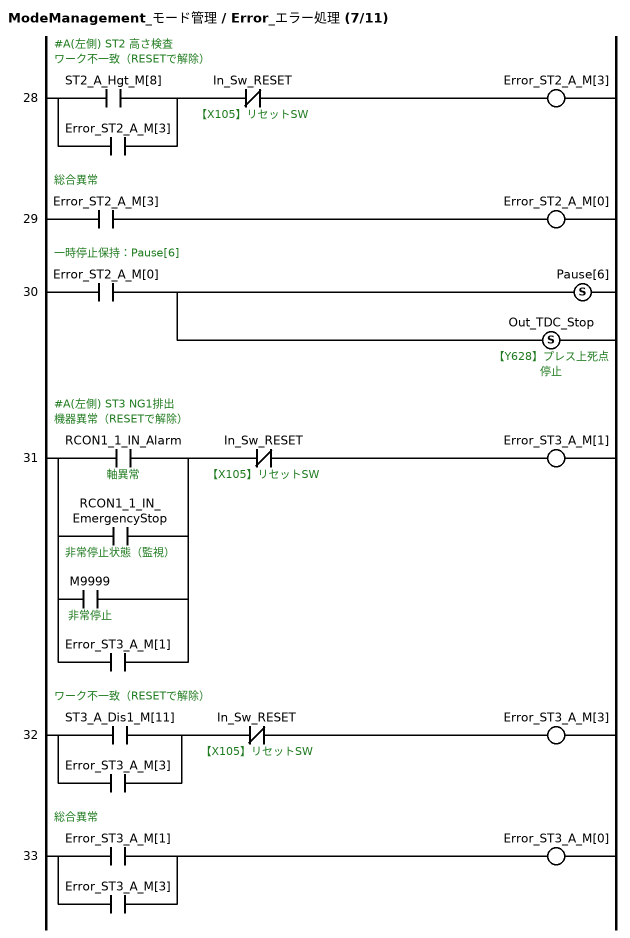
(* Rung 28: #A(左側) ST2 高さ検査 / ワーク不一致（RESETで解除） *)
Error_ST2_A_M[3] := (ST2_A_Hgt_M[8] OR Error_ST2_A_M[3]) AND NOT In_Sw_RESET;
(* Rung 29: 総合異常 *)
Error_ST2_A_M[0] := Error_ST2_A_M[3];
(* Rung 30: 一時停止保持：Pause[6] *)
IF Error_ST2_A_M[0] THEN
    Pause[6] := TRUE;
    Out_TDC_Stop := TRUE;
END_IF;
(* Rung 31: #A(左側) ST3 NG1排出 / 機器異常（RESETで解除） *)
Error_ST3_A_M[1] := (RCON1_1_IN_Alarm OR RCON1_1_IN_EmergencyStop OR M9999 OR Error_ST3_A_M[1]) AND NOT In_Sw_RESET;
(* Rung 32: ワーク不一致（RESETで解除） *)
Error_ST3_A_M[3] := (ST3_A_Dis1_M[11] OR Error_ST3_A_M[3]) AND NOT In_Sw_RESET;
(* Rung 33: 総合異常 *)
Error_ST3_A_M[0] := Error_ST3_A_M[1] OR Error_ST3_A_M[3];

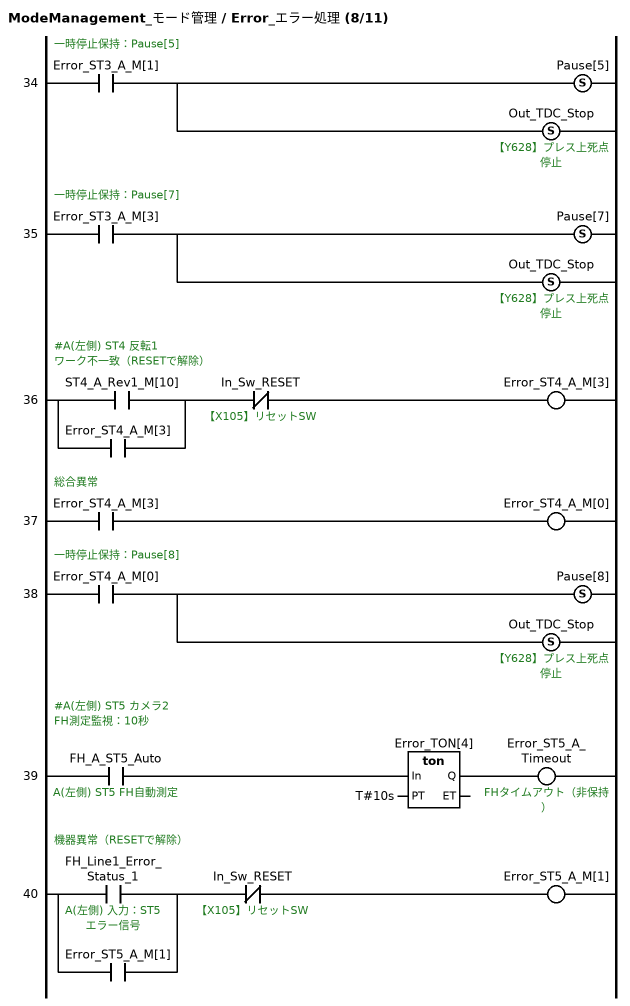
(* Rung 34: 一時停止保持：Pause[5] *)
IF Error_ST3_A_M[1] THEN
    Pause[5] := TRUE;
    Out_TDC_Stop := TRUE;
END_IF;
(* Rung 35: 一時停止保持：Pause[7] *)
IF Error_ST3_A_M[3] THEN
    Pause[7] := TRUE;
    Out_TDC_Stop := TRUE;
END_IF;
(* Rung 36: #A(左側) ST4 反転1 / ワーク不一致（RESETで解除） *)
Error_ST4_A_M[3] := (ST4_A_Rev1_M[10] OR Error_ST4_A_M[3]) AND NOT In_Sw_RESET;
(* Rung 37: 総合異常 *)
Error_ST4_A_M[0] := Error_ST4_A_M[3];
(* Rung 38: 一時停止保持：Pause[8] *)
IF Error_ST4_A_M[0] THEN
    Pause[8] := TRUE;
    Out_TDC_Stop := TRUE;
END_IF;
(* Rung 39: #A(左側) ST5 カメラ2 / FH測定監視：10秒 *)
Error_TON[4](In := FH_A_ST5_Auto, PT := T#10s);
Error_ST5_A_Timeout := Error_TON[4].Q;
(* Rung 40: 機器異常（RESETで解除） *)
Error_ST5_A_M[1] := (FH_Line1_Error_Status_1 OR Error_ST5_A_M[1]) AND NOT In_Sw_RESET;

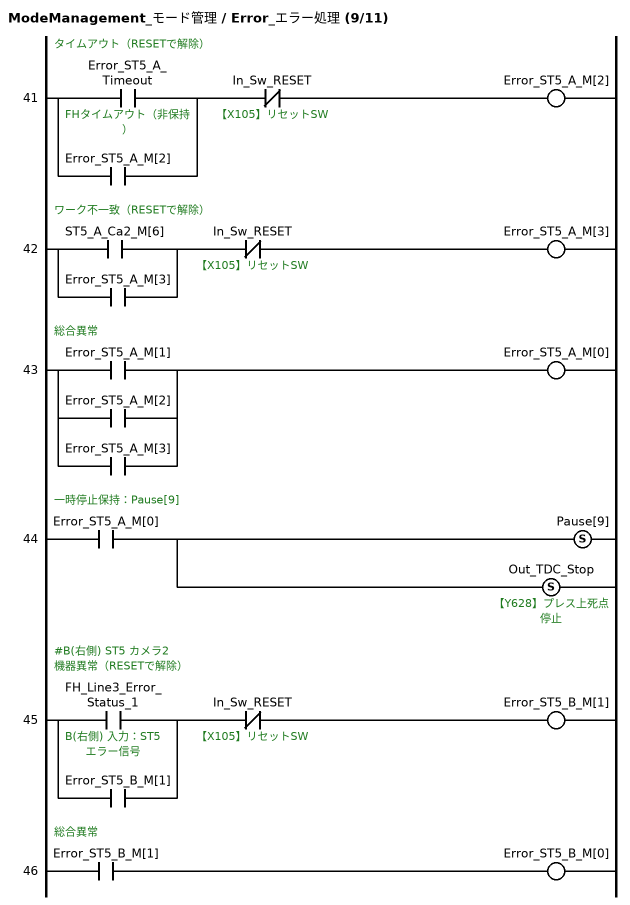
(* Rung 41: タイムアウト（RESETで解除） *)
Error_ST5_A_M[2] := (Error_ST5_A_Timeout OR Error_ST5_A_M[2]) AND NOT In_Sw_RESET;
(* Rung 42: ワーク不一致（RESETで解除） *)
Error_ST5_A_M[3] := (ST5_A_Ca2_M[6] OR Error_ST5_A_M[3]) AND NOT In_Sw_RESET;
(* Rung 43: 総合異常 *)
Error_ST5_A_M[0] := Error_ST5_A_M[1] OR Error_ST5_A_M[2] OR Error_ST5_A_M[3];
(* Rung 44: 一時停止保持：Pause[9] *)
IF Error_ST5_A_M[0] THEN
    Pause[9] := TRUE;
    Out_TDC_Stop := TRUE;
END_IF;
(* Rung 45: #B(右側) ST5 カメラ2 / 機器異常（RESETで解除） *)
Error_ST5_B_M[1] := (FH_Line3_Error_Status_1 OR Error_ST5_B_M[1]) AND NOT In_Sw_RESET;
(* Rung 46: 総合異常 *)
Error_ST5_B_M[0] := Error_ST5_B_M[1];

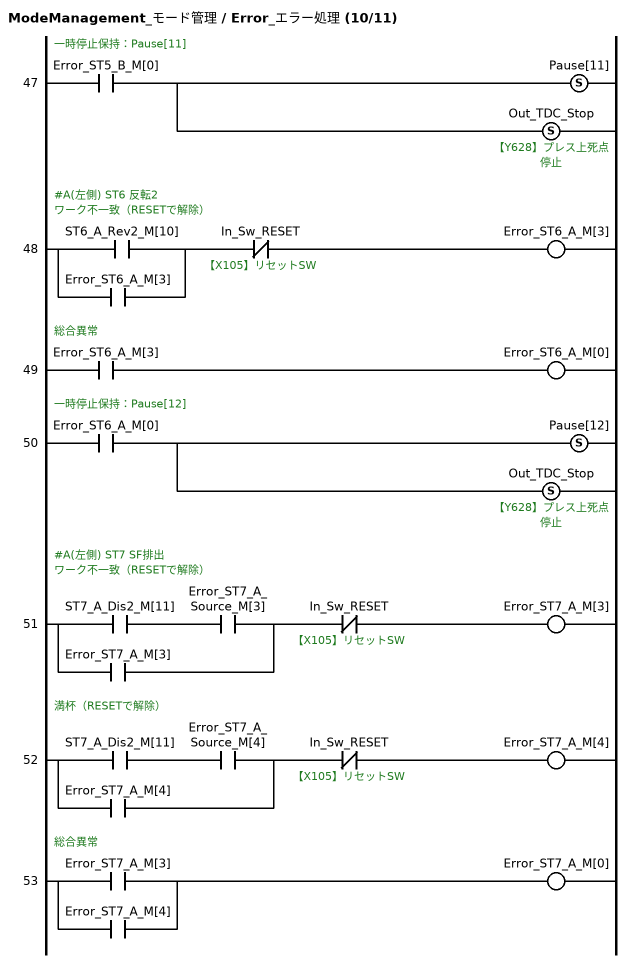
(* Rung 47: 一時停止保持：Pause[11] *)
IF Error_ST5_B_M[0] THEN
    Pause[11] := TRUE;
    Out_TDC_Stop := TRUE;
END_IF;
(* Rung 48: #A(左側) ST6 反転2 / ワーク不一致（RESETで解除） *)
Error_ST6_A_M[3] := (ST6_A_Rev2_M[10] OR Error_ST6_A_M[3]) AND NOT In_Sw_RESET;
(* Rung 49: 総合異常 *)
Error_ST6_A_M[0] := Error_ST6_A_M[3];
(* Rung 50: 一時停止保持：Pause[12] *)
IF Error_ST6_A_M[0] THEN
    Pause[12] := TRUE;
    Out_TDC_Stop := TRUE;
END_IF;
(* Rung 51: #A(左側) ST7 SF排出 / ワーク不一致（RESETで解除） *)
Error_ST7_A_M[3] := ((ST7_A_Dis2_M[11] AND Error_ST7_A_Source_M[3]) OR Error_ST7_A_M[3]) AND NOT In_Sw_RESET;
(* Rung 52: 満杯（RESETで解除） *)
Error_ST7_A_M[4] := ((ST7_A_Dis2_M[11] AND Error_ST7_A_Source_M[4]) OR Error_ST7_A_M[4]) AND NOT In_Sw_RESET;
(* Rung 53: 総合異常 *)
Error_ST7_A_M[0] := Error_ST7_A_M[3] OR Error_ST7_A_M[4];

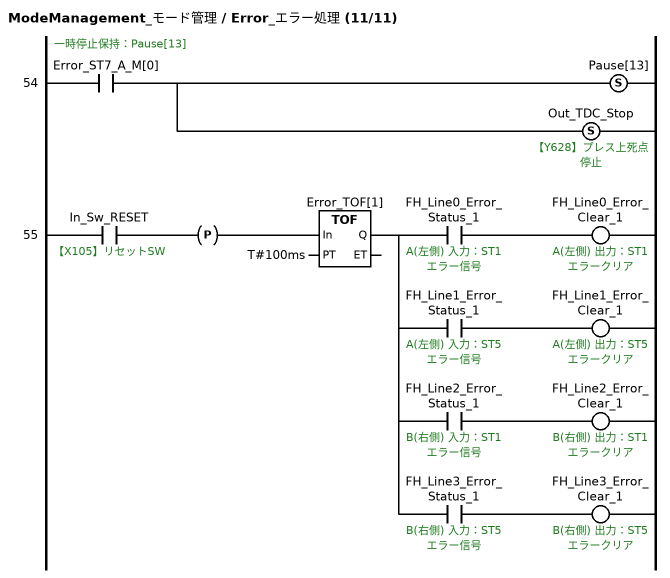
(* Rung 54: 一時停止保持：Pause[13] *)
IF Error_ST7_A_M[0] THEN
    Pause[13] := TRUE;
    Out_TDC_Stop := TRUE;
END_IF;
(* Rung 55 *)
_e45(CLK := In_Sw_RESET);
Error_TOF[1](In := _e45.Q, PT := T#100ms);
FH_Line0_Error_Clear_1 := Error_TOF[1].Q AND FH_Line0_Error_Status_1;
FH_Line1_Error_Clear_1 := Error_TOF[1].Q AND FH_Line1_Error_Status_1;
FH_Line2_Error_Clear_1 := Error_TOF[1].Q AND FH_Line2_Error_Status_1;
FH_Line3_Error_Clear_1 := Error_TOF[1].Q AND FH_Line3_Error_Status_1;

(* Section HMI_Request_表示要求: ladder, written here as Structured Text *)

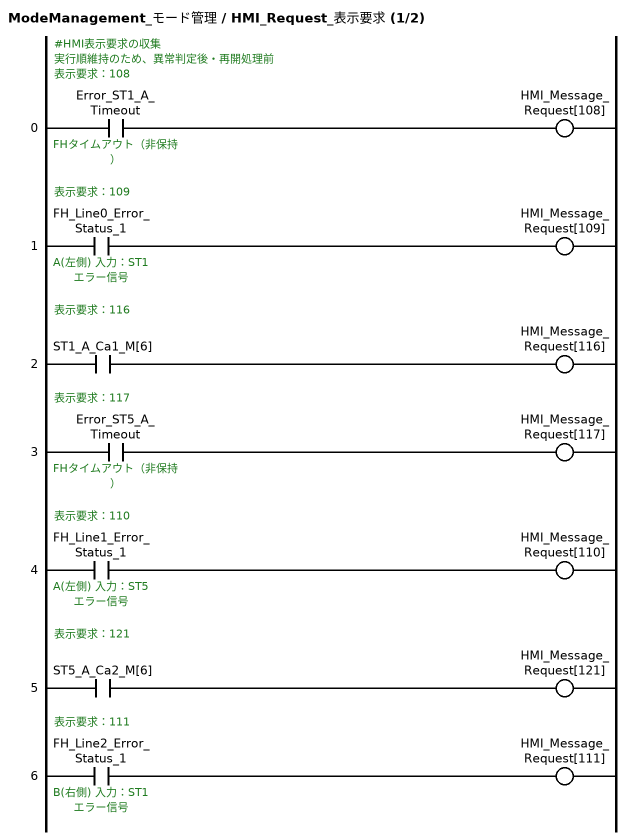
(* Rung 0: #HMI表示要求の収集 / 実行順維持のため、異常判定後・再開処理前 / 表示要求：108 *)
HMI_Message_Request[108] := Error_ST1_A_Timeout;
(* Rung 1: 表示要求：109 *)
HMI_Message_Request[109] := FH_Line0_Error_Status_1;
(* Rung 2: 表示要求：116 *)
HMI_Message_Request[116] := ST1_A_Ca1_M[6];
(* Rung 3: 表示要求：117 *)
HMI_Message_Request[117] := Error_ST5_A_Timeout;
(* Rung 4: 表示要求：110 *)
HMI_Message_Request[110] := FH_Line1_Error_Status_1;
(* Rung 5: 表示要求：121 *)
HMI_Message_Request[121] := ST5_A_Ca2_M[6];
(* Rung 6: 表示要求：111 *)
HMI_Message_Request[111] := FH_Line2_Error_Status_1;

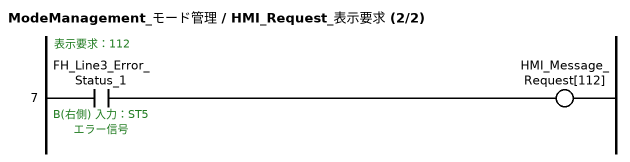
(* Rung 7: 表示要求：112 *)
HMI_Message_Request[112] := FH_Line3_Error_Status_1;

(* Section Restart_再開処理: ladder, written here as Structured Text *)

